REGION Network 1: จัดเก็บ
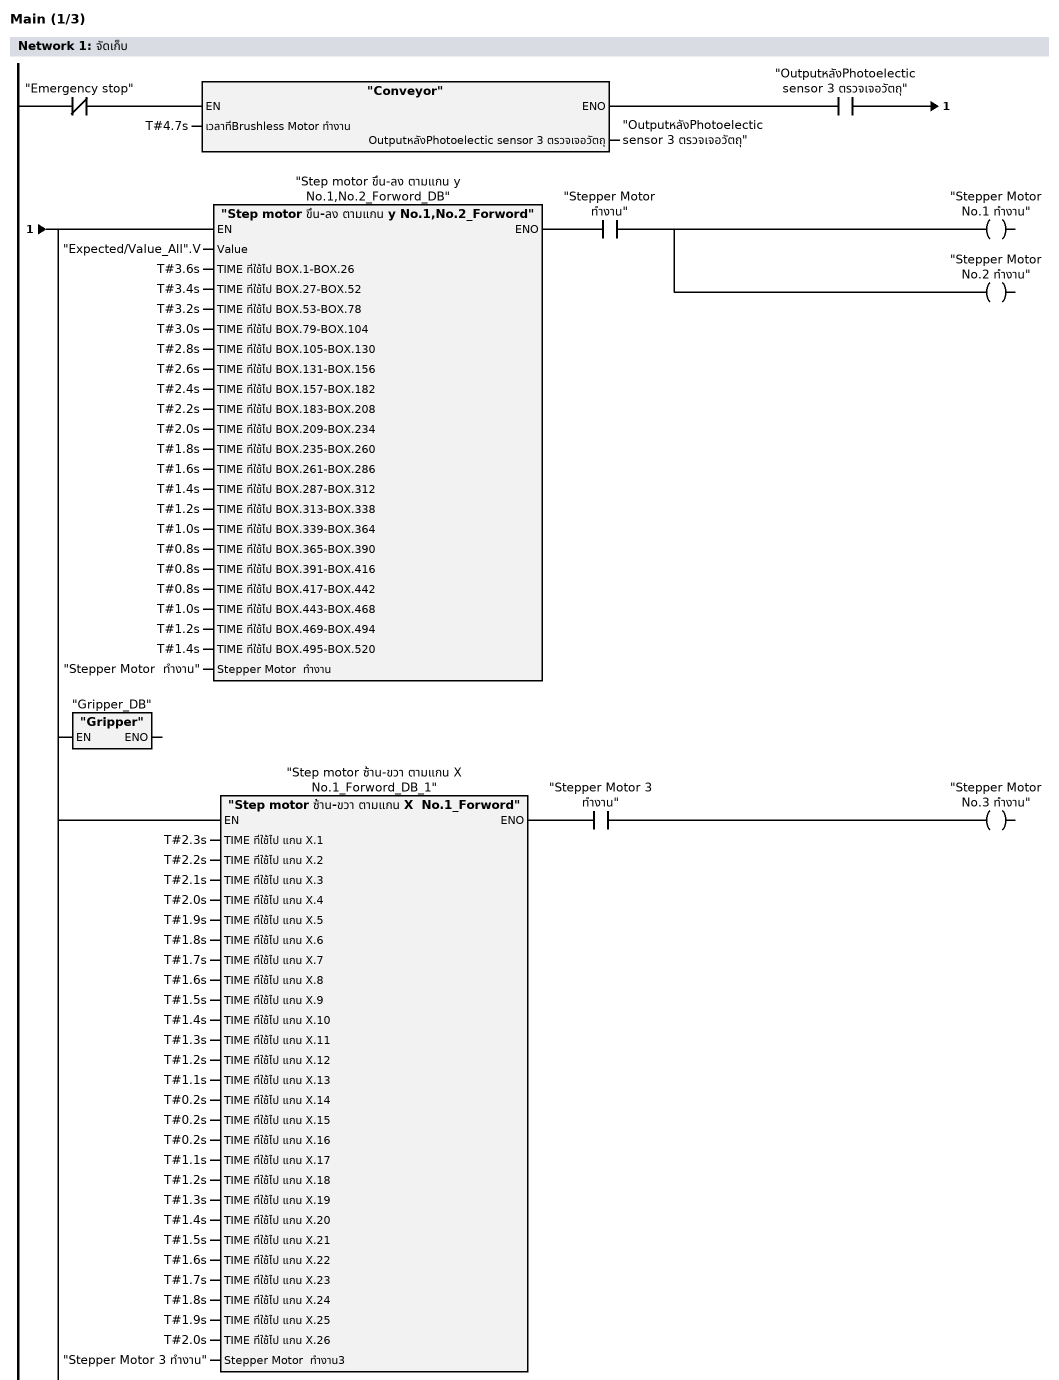
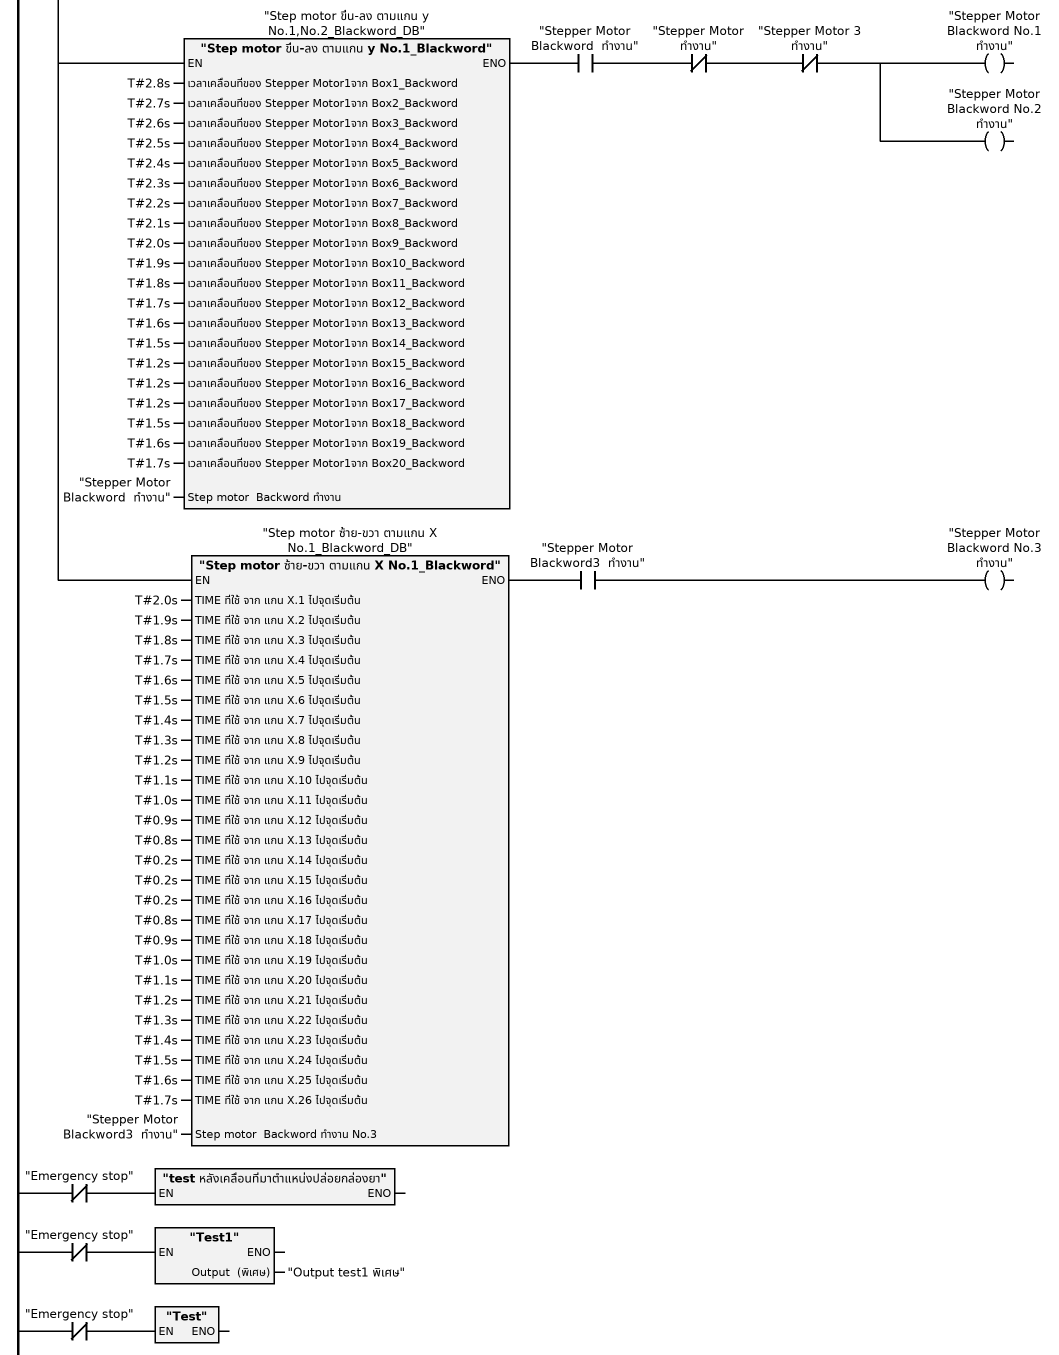
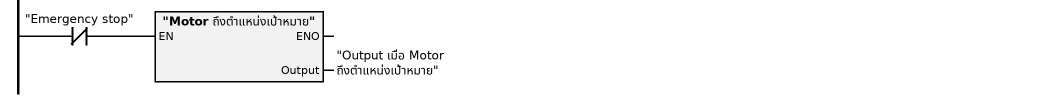
   RUNG wire#powerrail
      I_Contact( "Emergency stop" )
      "Conveyor"("เวลาที่Brushless Motor ทำงาน" := T#4.7s, "OutputหลังPhotoelectic sensor 3 ตรวจเจอวัตถุ" => "OutputหลังPhotoelectic sensor 3 ตรวจเจอวัตถุ")
      Contact( "OutputหลังPhotoelectic sensor 3 ตรวจเจอวัตถุ" )
      wire#w1
      "Step motor ขึ่น-ลง ตามแกน y No.1,No.2_Forword_DB"(Value := "Expected/Value_All".V, "TIME ที่ใช้ไป BOX.1-BOX.26" := T#3.6s, "TIME ที่ใช้ไป BOX.27-BOX.52" := T#3.4s, "TIME ที่ใช้ไป BOX.53-BOX.78" := T#3.2s, "TIME ที่ใช้ไป BOX.79-BOX.104" := T#3.0s, "TIME ที่ใช้ไป BOX.105-BOX.130" := T#2.8s, "TIME ที่ใช้ไป BOX.131-BOX.156" := T#2.6s, "TIME ที่ใช้ไป BOX.157-BOX.182" := T#2.4s, "TIME ที่ใช้ไป BOX.183-BOX.208" := T#2.2s, "TIME ที่ใช้ไป BOX.209-BOX.234" := T#2.0s, "TIME ที่ใช้ไป BOX.235-BOX.260" := T#1.8s, "TIME ที่ใช้ไป BOX.261-BOX.286" := T#1.6s, "TIME ที่ใช้ไป BOX.287-BOX.312" := T#1.4s, "TIME ที่ใช้ไป BOX.313-BOX.338" := T#1.2s, "TIME ที่ใช้ไป BOX.339-BOX.364" := T#1.0s, "TIME ที่ใช้ไป BOX.365-BOX.390" := T#0.8s, "TIME ที่ใช้ไป BOX.391-BOX.416" := T#0.8s, "TIME ที่ใช้ไป BOX.417-BOX.442" := T#0.8s, "TIME ที่ใช้ไป BOX.443-BOX.468" := T#1.0s, "TIME ที่ใช้ไป BOX.469-BOX.494" := T#1.2s, "TIME ที่ใช้ไป BOX.495-BOX.520" := T#1.4s, "Stepper Motor  ทำงาน" := "Stepper Motor  ทำงาน")
      Contact( "Stepper Motor  ทำงาน" )
      wire#w2
      Coil( "Stepper Motor No.1 ทำงาน" )
   END_RUNG
   RUNG wire#w2
      Coil( "Stepper Motor No.2 ทำงาน" )
   END_RUNG
   RUNG wire#w1
      "Gripper_DB"()
   END_RUNG
   RUNG wire#w1
      "Step motor ซ้าน-ขวา ตามแกน X  No.1_Forword_DB_1"("TIME ที่ใช้ไป แกน X.1" := T#2.3s, "TIME ที่ใช้ไป แกน X.2" := T#2.2s, "TIME ที่ใช้ไป แกน X.3" := T#2.1s, "TIME ที่ใช้ไป แกน X.4" := T#2.0s, "TIME ที่ใช้ไป แกน X.5" := T#1.9s, "TIME ที่ใช้ไป แกน X.6" := T#1.8s, "TIME ที่ใช้ไป แกน X.7" := T#1.7s, "TIME ที่ใช้ไป แกน X.8" := T#1.6s, "TIME ที่ใช้ไป แกน X.9" := T#1.5s, "TIME ที่ใช้ไป แกน X.10" := T#1.4s, "TIME ที่ใช้ไป แกน X.11" := T#1.3s, "TIME ที่ใช้ไป แกน X.12" := T#1.2s, "TIME ที่ใช้ไป แกน X.13" := T#1.1s, "TIME ที่ใช้ไป แกน X.14" := T#0.2s, "TIME ที่ใช้ไป แกน X.15" := T#0.2s, "TIME ที่ใช้ไป แกน X.16" := T#0.2s, "TIME ที่ใช้ไป แกน X.17" := T#1.1s, "TIME ที่ใช้ไป แกน X.18" := T#1.2s, "TIME ที่ใช้ไป แกน X.19" := T#1.3s, "TIME ที่ใช้ไป แกน X.20" := T#1.4s, "TIME ที่ใช้ไป แกน X.21" := T#1.5s, "TIME ที่ใช้ไป แกน X.22" := T#1.6s, "TIME ที่ใช้ไป แกน X.23" := T#1.7s, "TIME ที่ใช้ไป แกน X.24" := T#1.8s, "TIME ที่ใช้ไป แกน X.25" := T#1.9s, "TIME ที่ใช้ไป แกน X.26" := T#2.0s, "Stepper Motor  ทำงาน3" := "Stepper Motor 3 ทำงาน")
      Contact( "Stepper Motor 3 ทำงาน" )
      Coil( "Stepper Motor No.3 ทำงาน" )
   END_RUNG
   RUNG wire#w1
      "Step motor ขึ่น-ลง ตามแกน y No.1,No.2_Blackword_DB"("เวลาเคลื่อนที่ของ Stepper Motor1จาก Box1_Backword" := T#2.8s, "เวลาเคลื่อนที่ของ Stepper Motor1จาก Box2_Backword" := T#2.7s, "เวลาเคลื่อนที่ของ Stepper Motor1จาก Box3_Backword" := T#2.6s, "เวลาเคลื่อนที่ของ Stepper Motor1จาก Box4_Backword" := T#2.5s, "เวลาเคลื่อนที่ของ Stepper Motor1จาก Box5_Backword" := T#2.4s, "เวลาเคลื่อนที่ของ Stepper Motor1จาก Box6_Backword" := T#2.3s, "เวลาเคลื่อนที่ของ Stepper Motor1จาก Box7_Backword" := T#2.2s, "เวลาเคลื่อนที่ของ Stepper Motor1จาก Box8_Backword" := T#2.1s, "เวลาเคลื่อนที่ของ Stepper Motor1จาก Box9_Backword" := T#2.0s, "เวลาเคลื่อนที่ของ Stepper Motor1จาก Box10_Backword" := T#1.9s, "เวลาเคลื่อนที่ของ Stepper Motor1จาก Box11_Backword" := T#1.8s, "เวลาเคลื่อนที่ของ Stepper Motor1จาก Box12_Backword" := T#1.7s, "เวลาเคลื่อนที่ของ Stepper Motor1จาก Box13_Backword" := T#1.6s, "เวลาเคลื่อนที่ของ Stepper Motor1จาก Box14_Backword" := T#1.5s, "เวลาเคลื่อนที่ของ Stepper Motor1จาก Box15_Backword" := T#1.2s, "เวลาเคลื่อนที่ของ Stepper Motor1จาก Box16_Backword" := T#1.2s, "เวลาเคลื่อนที่ของ Stepper Motor1จาก Box17_Backword" := T#1.2s, "เวลาเคลื่อนที่ของ Stepper Motor1จาก Box18_Backword" := T#1.5s, "เวลาเคลื่อนที่ของ Stepper Motor1จาก Box19_Backword" := T#1.6s, "เวลาเคลื่อนที่ของ Stepper Motor1จาก Box20_Backword" := T#1.7s, "Step motor  Backword ทำงาน" := "Stepper Motor Blackword  ทำงาน")
      Contact( "Stepper Motor Blackword  ทำงาน" )
      I_Contact( "Stepper Motor  ทำงาน" )
      I_Contact( "Stepper Motor 3 ทำงาน" )
      wire#w3
      Coil( "Stepper Motor Blackword No.1 ทำงาน" )
   END_RUNG
   RUNG wire#w3
      Coil( "Stepper Motor Blackword No.2 ทำงาน" )
   END_RUNG
   RUNG wire#w1
      "Step motor ซ้าย-ขวา ตามแกน X No.1_Blackword_DB"("TIME ที่ใช้ จาก แกน X.1 ไปจุดเริ่มต้น" := T#2.0s, "TIME ที่ใช้ จาก แกน X.2 ไปจุดเริ่มต้น" := T#1.9s, "TIME ที่ใช้ จาก แกน X.3 ไปจุดเริ่มต้น" := T#1.8s, "TIME ที่ใช้ จาก แกน X.4 ไปจุดเริ่มต้น" := T#1.7s, "TIME ที่ใช้ จาก แกน X.5 ไปจุดเริ่มต้น" := T#1.6s, "TIME ที่ใช้ จาก แกน X.6 ไปจุดเริ่มต้น" := T#1.5s, "TIME ที่ใช้ จาก แกน X.7 ไปจุดเริ่มต้น" := T#1.4s, "TIME ที่ใช้ จาก แกน X.8 ไปจุดเริ่มต้น" := T#1.3s, "TIME ที่ใช้ จาก แกน X.9 ไปจุดเริ่มต้น" := T#1.2s, "TIME ที่ใช้ จาก แกน X.10 ไปจุดเริ่มต้น" := T#1.1s, "TIME ที่ใช้ จาก แกน X.11 ไปจุดเริ่มต้น" := T#1.0s, "TIME ที่ใช้ จาก แกน X.12 ไปจุดเริ่มต้น" := T#0.9s, "TIME ที่ใช้ จาก แกน X.13 ไปจุดเริ่มต้น" := T#0.8s, "TIME ที่ใช้ จาก แกน X.14 ไปจุดเริ่มต้น" := T#0.2s, "TIME ที่ใช้ จาก แกน X.15 ไปจุดเริ่มต้น" := T#0.2s, "TIME ที่ใช้ จาก แกน X.16 ไปจุดเริ่มต้น" := T#0.2s, "TIME ที่ใช้ จาก แกน X.17 ไปจุดเริ่มต้น" := T#0.8s, "TIME ที่ใช้ จาก แกน X.18 ไปจุดเริ่มต้น" := T#0.9s, "TIME ที่ใช้ จาก แกน X.19 ไปจุดเริ่มต้น" := T#1.0s, "TIME ที่ใช้ จาก แกน X.20 ไปจุดเริ่มต้น" := T#1.1s, "TIME ที่ใช้ จาก แกน X.21 ไปจุดเริ่มต้น" := T#1.2s, "TIME ที่ใช้ จาก แกน X.22 ไปจุดเริ่มต้น" := T#1.3s, "TIME ที่ใช้ จาก แกน X.23 ไปจุดเริ่มต้น" := T#1.4s, "TIME ที่ใช้ จาก แกน X.24 ไปจุดเริ่มต้น" := T#1.5s, "TIME ที่ใช้ จาก แกน X.25 ไปจุดเริ่มต้น" := T#1.6s, "TIME ที่ใช้ จาก แกน X.26 ไปจุดเริ่มต้น" := T#1.7s, "Step motor  Backword ทำงาน No.3" := "Stepper Motor Blackword3  ทำงาน")
      Contact( "Stepper Motor Blackword3  ทำงาน" )
      Coil( "Stepper Motor Blackword No.3 ทำงาน" )
   END_RUNG
   RUNG wire#powerrail
      I_Contact( "Emergency stop" )
      "test หลังเคลื่อนที่มาตำแหน่งปล่อยกล่องยา"()
   END_RUNG
   RUNG wire#powerrail
      I_Contact( "Emergency stop" )
      "Test1"("Output  (พิเศษ)" => "Output test1 พิเศษ")
   END_RUNG
   RUNG wire#powerrail
      I_Contact( "Emergency stop" )
      "Test"()
   END_RUNG
   RUNG wire#powerrail
      I_Contact( "Emergency stop" )
      "Motor ถึงตำแหน่งเป้าหมาย"(Output => "Output เมื่อ Motor ถึงตำแหน่งเป้าหมาย")
   END_RUNG
   // the same network as SCL:
   "Conveyor"(EN := NOT "Emergency stop",
              "เวลาที่Brushless Motor ทำงาน" := T#4.7s,
              "OutputหลังPhotoelectic sensor 3 ตรวจเจอวัตถุ" => "OutputหลังPhotoelectic sensor 3 ตรวจเจอวัตถุ",
              ENO => #_w1);
   #_w3 := #_w1 AND "OutputหลังPhotoelectic sensor 3 ตรวจเจอวัตถุ";
   "Step motor ขึ่น-ลง ตามแกน y No.1,No.2_Forword_DB"(EN := #_w1 AND "OutputหลังPhotoelectic sensor 3 ตรวจเจอวัตถุ",   // "Step motor ขึ่น-ลง ตามแกน y No.1,No.2_Forword"
                           Value := "Expected/Value_All".V,
                           "TIME ที่ใช้ไป BOX.1-BOX.26" := T#3.6s,
                           "TIME ที่ใช้ไป BOX.27-BOX.52" := T#3.4s,
                           "TIME ที่ใช้ไป BOX.53-BOX.78" := T#3.2s,
                           "TIME ที่ใช้ไป BOX.79-BOX.104" := T#3.0s,
                           "TIME ที่ใช้ไป BOX.105-BOX.130" := T#2.8s,
                           "TIME ที่ใช้ไป BOX.131-BOX.156" := T#2.6s,
                           "TIME ที่ใช้ไป BOX.157-BOX.182" := T#2.4s,
                           "TIME ที่ใช้ไป BOX.183-BOX.208" := T#2.2s,
                           "TIME ที่ใช้ไป BOX.209-BOX.234" := T#2.0s,
                           "TIME ที่ใช้ไป BOX.235-BOX.260" := T#1.8s,
                           "TIME ที่ใช้ไป BOX.261-BOX.286" := T#1.6s,
                           "TIME ที่ใช้ไป BOX.287-BOX.312" := T#1.4s,
                           "TIME ที่ใช้ไป BOX.313-BOX.338" := T#1.2s,
                           "TIME ที่ใช้ไป BOX.339-BOX.364" := T#1.0s,
                           "TIME ที่ใช้ไป BOX.365-BOX.390" := T#0.8s,
                           "TIME ที่ใช้ไป BOX.391-BOX.416" := T#0.8s,
                           "TIME ที่ใช้ไป BOX.417-BOX.442" := T#0.8s,
                           "TIME ที่ใช้ไป BOX.443-BOX.468" := T#1.0s,
                           "TIME ที่ใช้ไป BOX.469-BOX.494" := T#1.2s,
                           "TIME ที่ใช้ไป BOX.495-BOX.520" := T#1.4s,
                           "Stepper Motor  ทำงาน" := "Stepper Motor  ทำงาน",
                           ENO => #_w2);
   "Stepper Motor No.1 ทำงาน" := #_w2 AND "Stepper Motor  ทำงาน";
   "Stepper Motor No.2 ทำงาน" := "Stepper Motor No.1 ทำงาน";
   IF #_w3 THEN
       "Gripper_DB"();   // "Gripper"
   END_IF;
   "Step motor ซ้าน-ขวา ตามแกน X  No.1_Forword_DB_1"(EN := #_w3,   // "Step motor ซ้าน-ขวา ตามแกน X  No.1_Forword"
                           "TIME ที่ใช้ไป แกน X.1" := T#2.3s,
                           "TIME ที่ใช้ไป แกน X.2" := T#2.2s,
                           "TIME ที่ใช้ไป แกน X.3" := T#2.1s,
                           "TIME ที่ใช้ไป แกน X.4" := T#2.0s,
                           "TIME ที่ใช้ไป แกน X.5" := T#1.9s,
                           "TIME ที่ใช้ไป แกน X.6" := T#1.8s,
                           "TIME ที่ใช้ไป แกน X.7" := T#1.7s,
                           "TIME ที่ใช้ไป แกน X.8" := T#1.6s,
                           "TIME ที่ใช้ไป แกน X.9" := T#1.5s,
                           "TIME ที่ใช้ไป แกน X.10" := T#1.4s,
                           "TIME ที่ใช้ไป แกน X.11" := T#1.3s,
                           "TIME ที่ใช้ไป แกน X.12" := T#1.2s,
                           "TIME ที่ใช้ไป แกน X.13" := T#1.1s,
                           "TIME ที่ใช้ไป แกน X.14" := T#0.2s,
                           "TIME ที่ใช้ไป แกน X.15" := T#0.2s,
                           "TIME ที่ใช้ไป แกน X.16" := T#0.2s,
                           "TIME ที่ใช้ไป แกน X.17" := T#1.1s,
                           "TIME ที่ใช้ไป แกน X.18" := T#1.2s,
                           "TIME ที่ใช้ไป แกน X.19" := T#1.3s,
                           "TIME ที่ใช้ไป แกน X.20" := T#1.4s,
                           "TIME ที่ใช้ไป แกน X.21" := T#1.5s,
                           "TIME ที่ใช้ไป แกน X.22" := T#1.6s,
                           "TIME ที่ใช้ไป แกน X.23" := T#1.7s,
                           "TIME ที่ใช้ไป แกน X.24" := T#1.8s,
                           "TIME ที่ใช้ไป แกน X.25" := T#1.9s,
                           "TIME ที่ใช้ไป แกน X.26" := T#2.0s,
                           "Stepper Motor  ทำงาน3" := "Stepper Motor 3 ทำงาน",
                           ENO => #_w4);
   "Stepper Motor No.3 ทำงาน" := #_w4 AND "Stepper Motor 3 ทำงาน";
   "Step motor ขึ่น-ลง ตามแกน y No.1,No.2_Blackword_DB"(EN := #_w3,   // "Step motor ขึ่น-ลง ตามแกน y No.1_Blackword"
                           "เวลาเคลื่อนที่ของ Stepper Motor1จาก Box1_Backword" := T#2.8s,
                           "เวลาเคลื่อนที่ของ Stepper Motor1จาก Box2_Backword" := T#2.7s,
                           "เวลาเคลื่อนที่ของ Stepper Motor1จาก Box3_Backword" := T#2.6s,
                           "เวลาเคลื่อนที่ของ Stepper Motor1จาก Box4_Backword" := T#2.5s,
                           "เวลาเคลื่อนที่ของ Stepper Motor1จาก Box5_Backword" := T#2.4s,
                           "เวลาเคลื่อนที่ของ Stepper Motor1จาก Box6_Backword" := T#2.3s,
                           "เวลาเคลื่อนที่ของ Stepper Motor1จาก Box7_Backword" := T#2.2s,
                           "เวลาเคลื่อนที่ของ Stepper Motor1จาก Box8_Backword" := T#2.1s,
                           "เวลาเคลื่อนที่ของ Stepper Motor1จาก Box9_Backword" := T#2.0s,
                           "เวลาเคลื่อนที่ของ Stepper Motor1จาก Box10_Backword" := T#1.9s,
                           "เวลาเคลื่อนที่ของ Stepper Motor1จาก Box11_Backword" := T#1.8s,
                           "เวลาเคลื่อนที่ของ Stepper Motor1จาก Box12_Backword" := T#1.7s,
                           "เวลาเคลื่อนที่ของ Stepper Motor1จาก Box13_Backword" := T#1.6s,
                           "เวลาเคลื่อนที่ของ Stepper Motor1จาก Box14_Backword" := T#1.5s,
                           "เวลาเคลื่อนที่ของ Stepper Motor1จาก Box15_Backword" := T#1.2s,
                           "เวลาเคลื่อนที่ของ Stepper Motor1จาก Box16_Backword" := T#1.2s,
                           "เวลาเคลื่อนที่ของ Stepper Motor1จาก Box17_Backword" := T#1.2s,
                           "เวลาเคลื่อนที่ของ Stepper Motor1จาก Box18_Backword" := T#1.5s,
                           "เวลาเคลื่อนที่ของ Stepper Motor1จาก Box19_Backword" := T#1.6s,
                           "เวลาเคลื่อนที่ของ Stepper Motor1จาก Box20_Backword" := T#1.7s,
                           "Step motor  Backword ทำงาน" := "Stepper Motor Blackword  ทำงาน",
                           ENO => #_w5);
   "Stepper Motor Blackword No.1 ทำงาน" := #_w5 AND "Stepper Motor Blackword  ทำงาน" AND NOT "Stepper Motor  ทำงาน" AND NOT "Stepper Motor 3 ทำงาน";
   "Stepper Motor Blackword No.2 ทำงาน" := "Stepper Motor Blackword No.1 ทำงาน";
   "Step motor ซ้าย-ขวา ตามแกน X No.1_Blackword_DB"(EN := #_w3,   // "Step motor ซ้าย-ขวา ตามแกน X No.1_Blackword"
                           "TIME ที่ใช้ จาก แกน X.1 ไปจุดเริ่มต้น" := T#2.0s,
                           "TIME ที่ใช้ จาก แกน X.2 ไปจุดเริ่มต้น" := T#1.9s,
                           "TIME ที่ใช้ จาก แกน X.3 ไปจุดเริ่มต้น" := T#1.8s,
                           "TIME ที่ใช้ จาก แกน X.4 ไปจุดเริ่มต้น" := T#1.7s,
                           "TIME ที่ใช้ จาก แกน X.5 ไปจุดเริ่มต้น" := T#1.6s,
                           "TIME ที่ใช้ จาก แกน X.6 ไปจุดเริ่มต้น" := T#1.5s,
                           "TIME ที่ใช้ จาก แกน X.7 ไปจุดเริ่มต้น" := T#1.4s,
                           "TIME ที่ใช้ จาก แกน X.8 ไปจุดเริ่มต้น" := T#1.3s,
                           "TIME ที่ใช้ จาก แกน X.9 ไปจุดเริ่มต้น" := T#1.2s,
                           "TIME ที่ใช้ จาก แกน X.10 ไปจุดเริ่มต้น" := T#1.1s,
                           "TIME ที่ใช้ จาก แกน X.11 ไปจุดเริ่มต้น" := T#1.0s,
                           "TIME ที่ใช้ จาก แกน X.12 ไปจุดเริ่มต้น" := T#0.9s,
                           "TIME ที่ใช้ จาก แกน X.13 ไปจุดเริ่มต้น" := T#0.8s,
                           "TIME ที่ใช้ จาก แกน X.14 ไปจุดเริ่มต้น" := T#0.2s,
                           "TIME ที่ใช้ จาก แกน X.15 ไปจุดเริ่มต้น" := T#0.2s,
                           "TIME ที่ใช้ จาก แกน X.16 ไปจุดเริ่มต้น" := T#0.2s,
                           "TIME ที่ใช้ จาก แกน X.17 ไปจุดเริ่มต้น" := T#0.8s,
                           "TIME ที่ใช้ จาก แกน X.18 ไปจุดเริ่มต้น" := T#0.9s,
                           "TIME ที่ใช้ จาก แกน X.19 ไปจุดเริ่มต้น" := T#1.0s,
                           "TIME ที่ใช้ จาก แกน X.20 ไปจุดเริ่มต้น" := T#1.1s,
                           "TIME ที่ใช้ จาก แกน X.21 ไปจุดเริ่มต้น" := T#1.2s,
                           "TIME ที่ใช้ จาก แกน X.22 ไปจุดเริ่มต้น" := T#1.3s,
                           "TIME ที่ใช้ จาก แกน X.23 ไปจุดเริ่มต้น" := T#1.4s,
                           "TIME ที่ใช้ จาก แกน X.24 ไปจุดเริ่มต้น" := T#1.5s,
                           "TIME ที่ใช้ จาก แกน X.25 ไปจุดเริ่มต้น" := T#1.6s,
                           "TIME ที่ใช้ จาก แกน X.26 ไปจุดเริ่มต้น" := T#1.7s,
                           "Step motor  Backword ทำงาน No.3" := "Stepper Motor Blackword3  ทำงาน",
                           ENO => #_w6);
   "Stepper Motor Blackword No.3 ทำงาน" := #_w6 AND "Stepper Motor Blackword3  ทำงาน";
   IF NOT "Emergency stop" THEN "test หลังเคลื่อนที่มาตำแหน่งปล่อยกล่องยา"(); END_IF;
   IF NOT "Emergency stop" THEN "Test1"("Output  (พิเศษ)" => "Output test1 พิเศษ"); END_IF;
   IF NOT "Emergency stop" THEN "Test"(); END_IF;
   IF NOT "Emergency stop" THEN
       "Motor ถึงตำแหน่งเป้าหมาย"(Output => "Output เมื่อ Motor ถึงตำแหน่งเป้าหมาย");
   END_IF;
END_REGION

REGION Network 2: เบิกจ่าย
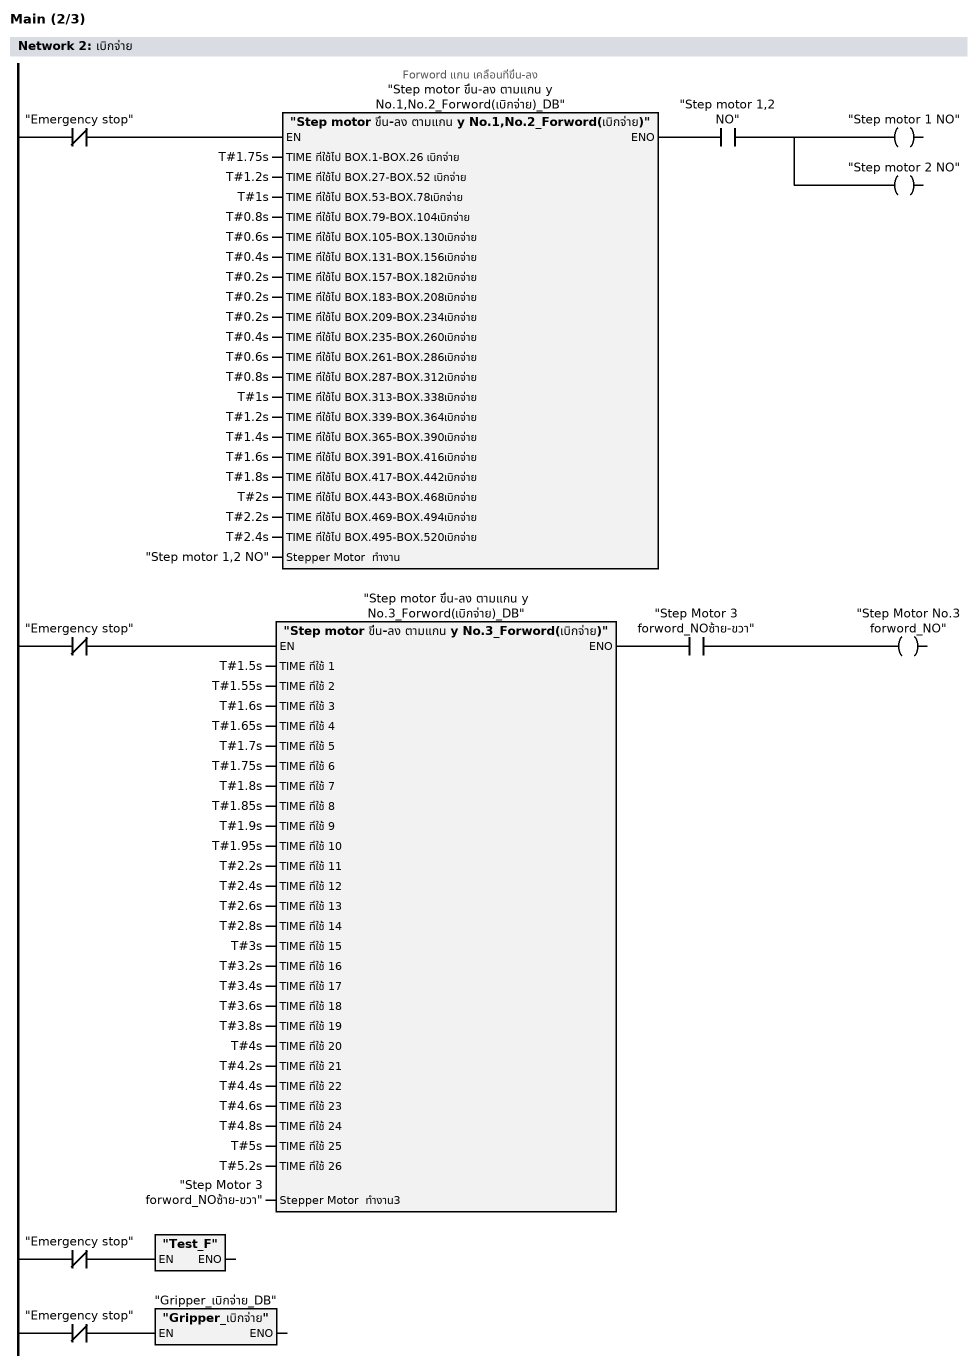
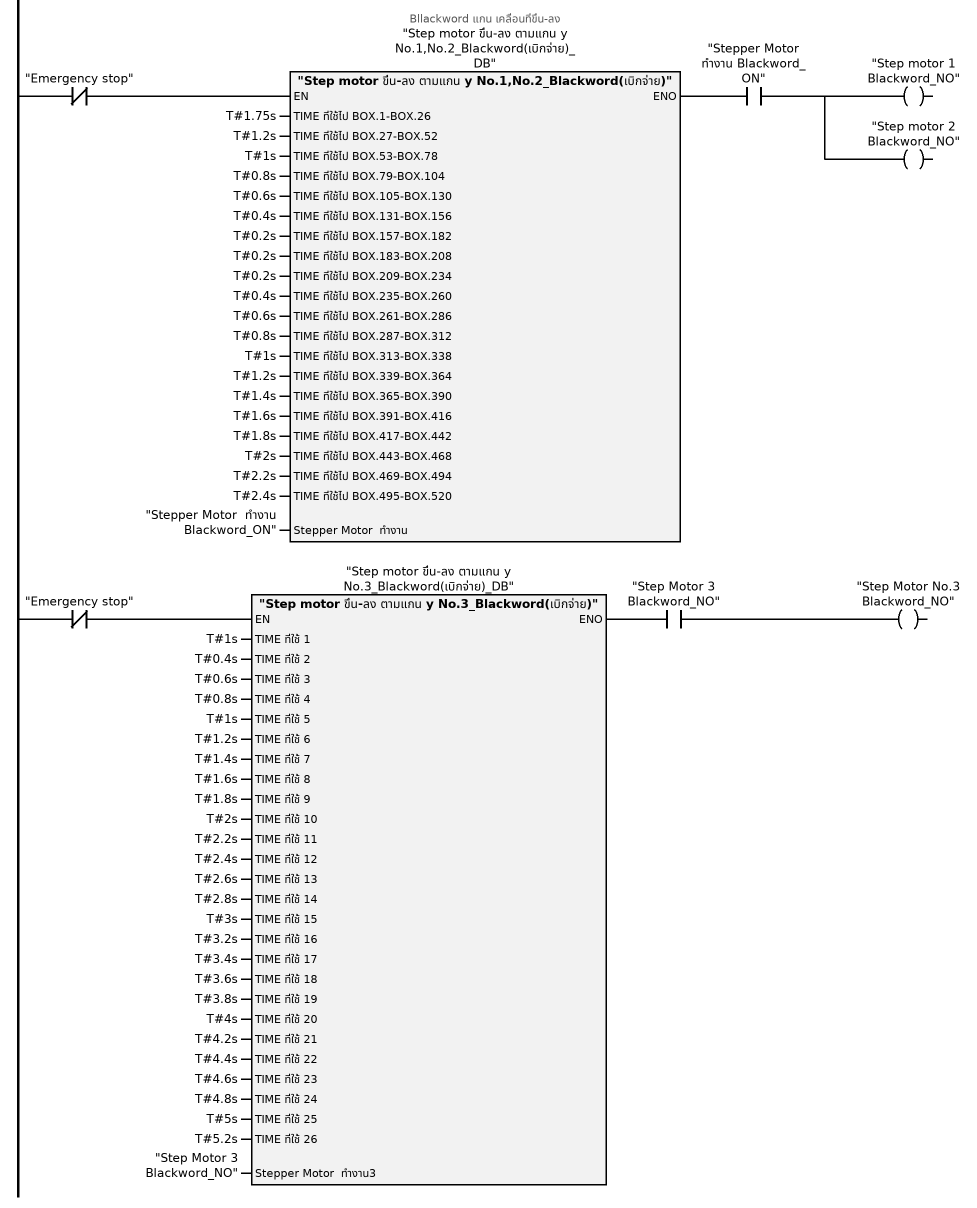
   RUNG wire#powerrail
      I_Contact( "Emergency stop" )
      "Step motor ขึ่น-ลง ตามแกน y No.1,No.2_Forword(เบิกจ่าย)_DB"("TIME ที่ใช้ไป BOX.1-BOX.26 เบิกจ่าย" := T#1.75s, "TIME ที่ใช้ไป BOX.27-BOX.52 เบิกจ่าย" := T#1.2s, "TIME ที่ใช้ไป BOX.53-BOX.78เบิกจ่าย" := T#1s, "TIME ที่ใช้ไป BOX.79-BOX.104เบิกจ่าย" := T#0.8s, "TIME ที่ใช้ไป BOX.105-BOX.130เบิกจ่าย" := T#0.6s, "TIME ที่ใช้ไป BOX.131-BOX.156เบิกจ่าย" := T#0.4s, "TIME ที่ใช้ไป BOX.157-BOX.182เบิกจ่าย" := T#0.2s, "TIME ที่ใช้ไป BOX.183-BOX.208เบิกจ่าย" := T#0.2s, "TIME ที่ใช้ไป BOX.209-BOX.234เบิกจ่าย" := T#0.2s, "TIME ที่ใช้ไป BOX.235-BOX.260เบิกจ่าย" := T#0.4s, "TIME ที่ใช้ไป BOX.261-BOX.286เบิกจ่าย" := T#0.6s, "TIME ที่ใช้ไป BOX.287-BOX.312เบิกจ่าย" := T#0.8s, "TIME ที่ใช้ไป BOX.313-BOX.338เบิกจ่าย" := T#1s, "TIME ที่ใช้ไป BOX.339-BOX.364เบิกจ่าย" := T#1.2s, "TIME ที่ใช้ไป BOX.365-BOX.390เบิกจ่าย" := T#1.4s, "TIME ที่ใช้ไป BOX.391-BOX.416เบิกจ่าย" := T#1.6s, "TIME ที่ใช้ไป BOX.417-BOX.442เบิกจ่าย" := T#1.8s, "TIME ที่ใช้ไป BOX.443-BOX.468เบิกจ่าย" := T#2s, "TIME ที่ใช้ไป BOX.469-BOX.494เบิกจ่าย" := T#2.2s, "TIME ที่ใช้ไป BOX.495-BOX.520เบิกจ่าย" := T#2.4s, "Stepper Motor  ทำงาน" := "Step motor 1,2 NO")   // Forword แกน เคลื่อนที่ขึ่น-ลง
      Contact( "Step motor 1,2 NO" )
      wire#w1
      Coil( "Step motor 1 NO" )
   END_RUNG
   RUNG wire#w1
      Coil( "Step motor 2 NO" )
   END_RUNG
   RUNG wire#powerrail
      I_Contact( "Emergency stop" )
      "Step motor ขึ่น-ลง ตามแกน y No.3_Forword(เบิกจ่าย)_DB"("TIME ที่ใช้ 1" := T#1.5s, "TIME ที่ใช้ 2" := T#1.55s, "TIME ที่ใช้ 3" := T#1.6s, "TIME ที่ใช้ 4" := T#1.65s, "TIME ที่ใช้ 5" := T#1.7s, "TIME ที่ใช้ 6" := T#1.75s, "TIME ที่ใช้ 7" := T#1.8s, "TIME ที่ใช้ 8" := T#1.85s, "TIME ที่ใช้ 9" := T#1.9s, "TIME ที่ใช้ 10" := T#1.95s, "TIME ที่ใช้ 11" := T#2.2s, "TIME ที่ใช้ 12" := T#2.4s, "TIME ที่ใช้ 13" := T#2.6s, "TIME ที่ใช้ 14" := T#2.8s, "TIME ที่ใช้ 15" := T#3s, "TIME ที่ใช้ 16" := T#3.2s, "TIME ที่ใช้ 17" := T#3.4s, "TIME ที่ใช้ 18" := T#3.6s, "TIME ที่ใช้ 19" := T#3.8s, "TIME ที่ใช้ 20" := T#4s, "TIME ที่ใช้ 21" := T#4.2s, "TIME ที่ใช้ 22" := T#4.4s, "TIME ที่ใช้ 23" := T#4.6s, "TIME ที่ใช้ 24" := T#4.8s, "TIME ที่ใช้ 25" := T#5s, "TIME ที่ใช้ 26" := T#5.2s, "Stepper Motor  ทำงาน3" := "Step Motor 3 forword_NOซ้าย-ขวา")
      Contact( "Step Motor 3 forword_NOซ้าย-ขวา" )
      Coil( "Step Motor No.3 forword_NO" )
   END_RUNG
   RUNG wire#powerrail
      I_Contact( "Emergency stop" )
      "Test_F"()
   END_RUNG
   RUNG wire#powerrail
      I_Contact( "Emergency stop" )
      "Gripper_เบิกจ่าย_DB"()
   END_RUNG
   RUNG wire#powerrail
      I_Contact( "Emergency stop" )
      "Step motor ขึ่น-ลง ตามแกน y No.1,No.2_Blackword(เบิกจ่าย)_DB"("TIME ที่ใช้ไป BOX.1-BOX.26" := T#1.75s, "TIME ที่ใช้ไป BOX.27-BOX.52" := T#1.2s, "TIME ที่ใช้ไป BOX.53-BOX.78" := T#1s, "TIME ที่ใช้ไป BOX.79-BOX.104" := T#0.8s, "TIME ที่ใช้ไป BOX.105-BOX.130" := T#0.6s, "TIME ที่ใช้ไป BOX.131-BOX.156" := T#0.4s, "TIME ที่ใช้ไป BOX.157-BOX.182" := T#0.2s, "TIME ที่ใช้ไป BOX.183-BOX.208" := T#0.2s, "TIME ที่ใช้ไป BOX.209-BOX.234" := T#0.2s, "TIME ที่ใช้ไป BOX.235-BOX.260" := T#0.4s, "TIME ที่ใช้ไป BOX.261-BOX.286" := T#0.6s, "TIME ที่ใช้ไป BOX.287-BOX.312" := T#0.8s, "TIME ที่ใช้ไป BOX.313-BOX.338" := T#1s, "TIME ที่ใช้ไป BOX.339-BOX.364" := T#1.2s, "TIME ที่ใช้ไป BOX.365-BOX.390" := T#1.4s, "TIME ที่ใช้ไป BOX.391-BOX.416" := T#1.6s, "TIME ที่ใช้ไป BOX.417-BOX.442" := T#1.8s, "TIME ที่ใช้ไป BOX.443-BOX.468" := T#2s, "TIME ที่ใช้ไป BOX.469-BOX.494" := T#2.2s, "TIME ที่ใช้ไป BOX.495-BOX.520" := T#2.4s, "Stepper Motor  ทำงาน" := "Stepper Motor  ทำงาน Blackword_ON")   // Bllackword แกน เคลื่อนที่ขึ่น-ลง
      Contact( "Stepper Motor  ทำงาน Blackword_ON" )
      wire#w2
      Coil( "Step motor 1 Blackword_NO" )
   END_RUNG
   RUNG wire#w2
      Coil( "Step motor 2 Blackword_NO" )
   END_RUNG
   RUNG wire#powerrail
      I_Contact( "Emergency stop" )
      "Step motor ขึ่น-ลง ตามแกน y No.3_Blackword(เบิกจ่าย)_DB"("TIME ที่ใช้ 1" := T#1s, "TIME ที่ใช้ 2" := T#0.4s, "TIME ที่ใช้ 3" := T#0.6s, "TIME ที่ใช้ 4" := T#0.8s, "TIME ที่ใช้ 5" := T#1s, "TIME ที่ใช้ 6" := T#1.2s, "TIME ที่ใช้ 7" := T#1.4s, "TIME ที่ใช้ 8" := T#1.6s, "TIME ที่ใช้ 9" := T#1.8s, "TIME ที่ใช้ 10" := T#2s, "TIME ที่ใช้ 11" := T#2.2s, "TIME ที่ใช้ 12" := T#2.4s, "TIME ที่ใช้ 13" := T#2.6s, "TIME ที่ใช้ 14" := T#2.8s, "TIME ที่ใช้ 15" := T#3s, "TIME ที่ใช้ 16" := T#3.2s, "TIME ที่ใช้ 17" := T#3.4s, "TIME ที่ใช้ 18" := T#3.6s, "TIME ที่ใช้ 19" := T#3.8s, "TIME ที่ใช้ 20" := T#4s, "TIME ที่ใช้ 21" := T#4.2s, "TIME ที่ใช้ 22" := T#4.4s, "TIME ที่ใช้ 23" := T#4.6s, "TIME ที่ใช้ 24" := T#4.8s, "TIME ที่ใช้ 25" := T#5s, "TIME ที่ใช้ 26" := T#5.2s, "Stepper Motor  ทำงาน3" := "Step Motor 3 Blackword_NO")
      Contact( "Step Motor 3 Blackword_NO" )
      Coil( "Step Motor No.3 Blackword_NO" )
   END_RUNG
   // the same network as SCL:
   "Step motor ขึ่น-ลง ตามแกน y No.1,No.2_Forword(เบิกจ่าย)_DB"(EN := NOT "Emergency stop",   // "Step motor ขึ่น-ลง ตามแกน y No.1,No.2_Forword(เบิกจ่าย)": Forword แกน เคลื่อนที่ขึ่น-ลง
                           "TIME ที่ใช้ไป BOX.1-BOX.26 เบิกจ่าย" := T#1.75s,
                           "TIME ที่ใช้ไป BOX.27-BOX.52 เบิกจ่าย" := T#1.2s,
                           "TIME ที่ใช้ไป BOX.53-BOX.78เบิกจ่าย" := T#1s,
                           "TIME ที่ใช้ไป BOX.79-BOX.104เบิกจ่าย" := T#0.8s,
                           "TIME ที่ใช้ไป BOX.105-BOX.130เบิกจ่าย" := T#0.6s,
                           "TIME ที่ใช้ไป BOX.131-BOX.156เบิกจ่าย" := T#0.4s,
                           "TIME ที่ใช้ไป BOX.157-BOX.182เบิกจ่าย" := T#0.2s,
                           "TIME ที่ใช้ไป BOX.183-BOX.208เบิกจ่าย" := T#0.2s,
                           "TIME ที่ใช้ไป BOX.209-BOX.234เบิกจ่าย" := T#0.2s,
                           "TIME ที่ใช้ไป BOX.235-BOX.260เบิกจ่าย" := T#0.4s,
                           "TIME ที่ใช้ไป BOX.261-BOX.286เบิกจ่าย" := T#0.6s,
                           "TIME ที่ใช้ไป BOX.287-BOX.312เบิกจ่าย" := T#0.8s,
                           "TIME ที่ใช้ไป BOX.313-BOX.338เบิกจ่าย" := T#1s,
                           "TIME ที่ใช้ไป BOX.339-BOX.364เบิกจ่าย" := T#1.2s,
                           "TIME ที่ใช้ไป BOX.365-BOX.390เบิกจ่าย" := T#1.4s,
                           "TIME ที่ใช้ไป BOX.391-BOX.416เบิกจ่าย" := T#1.6s,
                           "TIME ที่ใช้ไป BOX.417-BOX.442เบิกจ่าย" := T#1.8s,
                           "TIME ที่ใช้ไป BOX.443-BOX.468เบิกจ่าย" := T#2s,
                           "TIME ที่ใช้ไป BOX.469-BOX.494เบิกจ่าย" := T#2.2s,
                           "TIME ที่ใช้ไป BOX.495-BOX.520เบิกจ่าย" := T#2.4s,
                           "Stepper Motor  ทำงาน" := "Step motor 1,2 NO",
                           ENO => #_w1);
   "Step motor 1 NO" := #_w1 AND "Step motor 1,2 NO";
   "Step motor 2 NO" := "Step motor 1 NO";
   "Step motor ขึ่น-ลง ตามแกน y No.3_Forword(เบิกจ่าย)_DB"(EN := NOT "Emergency stop",   // "Step motor ขึ่น-ลง ตามแกน y No.3_Forword(เบิกจ่าย)"
                           "TIME ที่ใช้ 1" := T#1.5s,
                           "TIME ที่ใช้ 2" := T#1.55s,
                           "TIME ที่ใช้ 3" := T#1.6s,
                           "TIME ที่ใช้ 4" := T#1.65s,
                           "TIME ที่ใช้ 5" := T#1.7s,
                           "TIME ที่ใช้ 6" := T#1.75s,
                           "TIME ที่ใช้ 7" := T#1.8s,
                           "TIME ที่ใช้ 8" := T#1.85s,
                           "TIME ที่ใช้ 9" := T#1.9s,
                           "TIME ที่ใช้ 10" := T#1.95s,
                           "TIME ที่ใช้ 11" := T#2.2s,
                           "TIME ที่ใช้ 12" := T#2.4s,
                           "TIME ที่ใช้ 13" := T#2.6s,
                           "TIME ที่ใช้ 14" := T#2.8s,
                           "TIME ที่ใช้ 15" := T#3s,
                           "TIME ที่ใช้ 16" := T#3.2s,
                           "TIME ที่ใช้ 17" := T#3.4s,
                           "TIME ที่ใช้ 18" := T#3.6s,
                           "TIME ที่ใช้ 19" := T#3.8s,
                           "TIME ที่ใช้ 20" := T#4s,
                           "TIME ที่ใช้ 21" := T#4.2s,
                           "TIME ที่ใช้ 22" := T#4.4s,
                           "TIME ที่ใช้ 23" := T#4.6s,
                           "TIME ที่ใช้ 24" := T#4.8s,
                           "TIME ที่ใช้ 25" := T#5s,
                           "TIME ที่ใช้ 26" := T#5.2s,
                           "Stepper Motor  ทำงาน3" := "Step Motor 3 forword_NOซ้าย-ขวา",
                           ENO => #_w2);
   "Step Motor No.3 forword_NO" := #_w2 AND "Step Motor 3 forword_NOซ้าย-ขวา";
   IF NOT "Emergency stop" THEN "Test_F"(); END_IF;
   IF NOT "Emergency stop" THEN
       "Gripper_เบิกจ่าย_DB"();   // "Gripper_เบิกจ่าย"
   END_IF;
   "Step motor ขึ่น-ลง ตามแกน y No.1,No.2_Blackword(เบิกจ่าย)_DB"(EN := NOT "Emergency stop",   // "Step motor ขึ่น-ลง ตามแกน y No.1,No.2_Blackword(เบิกจ่าย)": Bllackword แกน เคลื่อนที่ขึ่น-ลง
                           "TIME ที่ใช้ไป BOX.1-BOX.26" := T#1.75s,
                           "TIME ที่ใช้ไป BOX.27-BOX.52" := T#1.2s,
                           "TIME ที่ใช้ไป BOX.53-BOX.78" := T#1s,
                           "TIME ที่ใช้ไป BOX.79-BOX.104" := T#0.8s,
                           "TIME ที่ใช้ไป BOX.105-BOX.130" := T#0.6s,
                           "TIME ที่ใช้ไป BOX.131-BOX.156" := T#0.4s,
                           "TIME ที่ใช้ไป BOX.157-BOX.182" := T#0.2s,
                           "TIME ที่ใช้ไป BOX.183-BOX.208" := T#0.2s,
                           "TIME ที่ใช้ไป BOX.209-BOX.234" := T#0.2s,
                           "TIME ที่ใช้ไป BOX.235-BOX.260" := T#0.4s,
                           "TIME ที่ใช้ไป BOX.261-BOX.286" := T#0.6s,
                           "TIME ที่ใช้ไป BOX.287-BOX.312" := T#0.8s,
                           "TIME ที่ใช้ไป BOX.313-BOX.338" := T#1s,
                           "TIME ที่ใช้ไป BOX.339-BOX.364" := T#1.2s,
                           "TIME ที่ใช้ไป BOX.365-BOX.390" := T#1.4s,
                           "TIME ที่ใช้ไป BOX.391-BOX.416" := T#1.6s,
                           "TIME ที่ใช้ไป BOX.417-BOX.442" := T#1.8s,
                           "TIME ที่ใช้ไป BOX.443-BOX.468" := T#2s,
                           "TIME ที่ใช้ไป BOX.469-BOX.494" := T#2.2s,
                           "TIME ที่ใช้ไป BOX.495-BOX.520" := T#2.4s,
                           "Stepper Motor  ทำงาน" := "Stepper Motor  ทำงาน Blackword_ON",
                           ENO => #_w3);
   "Step motor 1 Blackword_NO" := #_w3 AND "Stepper Motor  ทำงาน Blackword_ON";
   "Step motor 2 Blackword_NO" := "Step motor 1 Blackword_NO";
   "Step motor ขึ่น-ลง ตามแกน y No.3_Blackword(เบิกจ่าย)_DB"(EN := NOT "Emergency stop",   // "Step motor ขึ่น-ลง ตามแกน y No.3_Blackword(เบิกจ่าย)"
                           "TIME ที่ใช้ 1" := T#1s,
                           "TIME ที่ใช้ 2" := T#0.4s,
                           "TIME ที่ใช้ 3" := T#0.6s,
                           "TIME ที่ใช้ 4" := T#0.8s,
                           "TIME ที่ใช้ 5" := T#1s,
                           "TIME ที่ใช้ 6" := T#1.2s,
                           "TIME ที่ใช้ 7" := T#1.4s,
                           "TIME ที่ใช้ 8" := T#1.6s,
                           "TIME ที่ใช้ 9" := T#1.8s,
                           "TIME ที่ใช้ 10" := T#2s,
                           "TIME ที่ใช้ 11" := T#2.2s,
                           "TIME ที่ใช้ 12" := T#2.4s,
                           "TIME ที่ใช้ 13" := T#2.6s,
                           "TIME ที่ใช้ 14" := T#2.8s,
                           "TIME ที่ใช้ 15" := T#3s,
                           "TIME ที่ใช้ 16" := T#3.2s,
                           "TIME ที่ใช้ 17" := T#3.4s,
                           "TIME ที่ใช้ 18" := T#3.6s,
                           "TIME ที่ใช้ 19" := T#3.8s,
                           "TIME ที่ใช้ 20" := T#4s,
                           "TIME ที่ใช้ 21" := T#4.2s,
                           "TIME ที่ใช้ 22" := T#4.4s,
                           "TIME ที่ใช้ 23" := T#4.6s,
                           "TIME ที่ใช้ 24" := T#4.8s,
                           "TIME ที่ใช้ 25" := T#5s,
                           "TIME ที่ใช้ 26" := T#5.2s,
                           "Stepper Motor  ทำงาน3" := "Step Motor 3 Blackword_NO",
                           ENO => #_w4);
   "Step Motor No.3 Blackword_NO" := #_w4 AND "Step Motor 3 Blackword_NO";
END_REGION

REGION Network 3: Screen
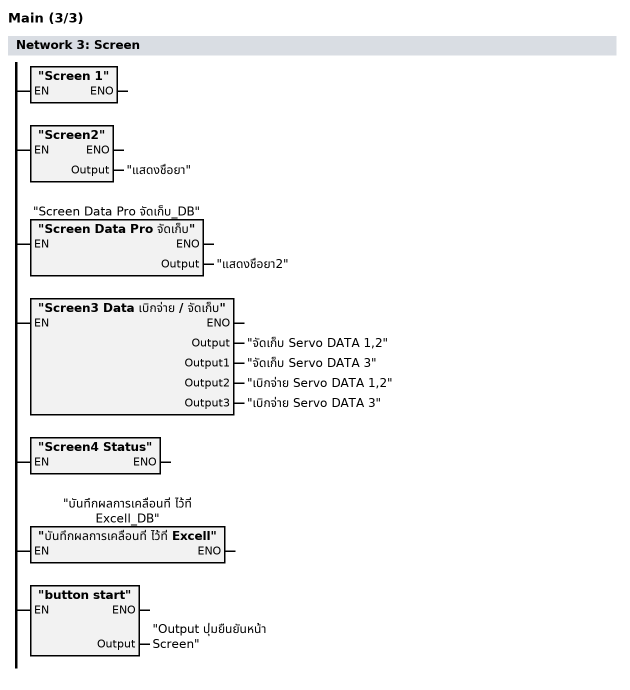
   RUNG wire#powerrail
      "Screen 1"()
   END_RUNG
   RUNG wire#powerrail
      "Screen2"(Output => "แสดงชื่อยา")
   END_RUNG
   RUNG wire#powerrail
      "Screen Data Pro จัดเก็บ_DB"(Output => "แสดงชื่อยา2")
   END_RUNG
   RUNG wire#powerrail
      "Screen3 Data เบิกจ่าย / จัดเก็บ"(Output => "จัดเก็บ Servo DATA 1,2", Output1 => "จัดเก็บ Servo DATA 3", Output2 => "เบิกจ่าย Servo DATA 1,2", Output3 => "เบิกจ่าย Servo DATA 3")
   END_RUNG
   RUNG wire#powerrail
      "Screen4 Status"()
   END_RUNG
   RUNG wire#powerrail
      "บันทึกผลการเคลื่อนที่ ไว้ที่ Excell_DB"()
   END_RUNG
   RUNG wire#powerrail
      "button start"(Output => "Output ปุ่มยืนยันหน้า Screen")
   END_RUNG
   // the same network as SCL:
   "Screen 1"();
   "Screen2"(Output => "แสดงชื่อยา");
   "Screen Data Pro จัดเก็บ_DB"(Output => "แสดงชื่อยา2");   // "Screen Data Pro จัดเก็บ"
   "Screen3 Data เบิกจ่าย / จัดเก็บ"(Output => "จัดเก็บ Servo DATA 1,2",
                           Output1 => "จัดเก็บ Servo DATA 3",
                           Output2 => "เบิกจ่าย Servo DATA 1,2",
                           Output3 => "เบิกจ่าย Servo DATA 3");
   "Screen4 Status"();
   "บันทึกผลการเคลื่อนที่ ไว้ที่ Excell_DB"();   // "บันทึกผลการเคลื่อนที่ ไว้ที่ Excell"
   "button start"(Output => "Output ปุ่มยืนยันหน้า Screen");
END_REGION
END_ORGANIZATION_BLOCK

// folder: GRAPH

FUNCTION_BLOCK "GRAPH_จัดเก็บ"   // FB17, GRAPH_PLUS
{ S7_Optimized_Access := 'TRUE' }
VERSION : 0.1
   VAR_INPUT
      OFF_SQ : Bool := false;   // Turn sequence off
      INIT_SQ : Bool := false;   // Set sequence to initial state
      ACK_EF : Bool := false;   // Acknowledge all errors and faults
      S_PREV : Bool := false;   // Output previous step in parameter S_NO
      S_NEXT : Bool := false;   // Indicate next step in parameter S_NO
      SW_AUTO : Bool := false;   // Automatic mode
      SW_TAP : Bool := false;   // Semiautomatic/switch with transition
      SW_TOP : Bool := false;   // Semiautomatic/ignore transition
      SW_MAN : Bool := false;   // Manual mode
      S_SEL : Int := 0;   // Select step to be output to S_NO
      S_ON : Bool := false;   // Activate step indicated in S_NO
      S_OFF : Bool := false;   // Deactivate step indicated S_NO
      T_PUSH : Bool := false;   // Enable transition to switch in semi automatic mode
   END_VAR
   VAR_OUTPUT
      S_NO : Int := 0;   // Step number
      S_MORE : Bool := false;   // More steps are available and can be shown in S_NO
      S_ACTIVE : Bool := false;   // Step indicated in S_NO is active
      ERR_FLT : Bool := false;   // Interlock or supervision group error
      AUTO_ON : Bool := false;   // Automatic mode is active
      TAP_ON : Bool := false;   // Semiautomatic mode/step with transition enabled
      TOP_ON : Bool := false;   // Semiautomatic mode/ignore transition enabled
      MAN_ON : Bool := false;   // Manual mode is active
   END_VAR
   VAR
      HMI_INFO : Array[0..8] of UInt;
      IF_PAR : G7_IfParPlus_V6;
      RT_DATA : G7_RTDataPlus_V6;   // Internal data area
      Trans1 : G7_TransitionPlus_V6;   // Transition structure
      Trans2 : G7_TransitionPlus_V6;   // Transition structure
      Trans3 : G7_TransitionPlus_V6;   // Transition structure
      Trans4 : G7_TransitionPlus_V6;   // Transition structure
      Trans5 : G7_TransitionPlus_V6;   // Transition structure
      Trans6 : G7_TransitionPlus_V6;   // Transition structure
      Trans7 : G7_TransitionPlus_V6;   // Transition structure
      Trans8 : G7_TransitionPlus_V6;   // Transition structure
      Trans9 : G7_TransitionPlus_V6;   // Transition structure
      Trans10 : G7_TransitionPlus_V6;   // Transition structure
      Trans11 : G7_TransitionPlus_V6;   // Transition structure
      Trans12 : G7_TransitionPlus_V6;   // Transition structure
      Trans13 : G7_TransitionPlus_V6;   // Transition structure
      Trans14 : G7_TransitionPlus_V6;   // Transition structure
      "รอรับคำสั่งยา" : G7_StepPlus_V6;   // Step structure
      "Conveyorลำเลียงกล่องยาไปตำแหน่งหยิบยา" : G7_StepPlus_V6;   // Step structure
      "หมุนไปจุดเริ่มต้น" : G7_StepPlus_V6;   // Step structure
      "gripper สไลด์ออกรับยา" : G7_StepPlus_V6;   // Step structure
      "gripper หนีบกล่องยา" : G7_StepPlus_V6;   // Step structure
      "gripper สไลด์เข้า" : G7_StepPlus_V6;   // Step structure
      "gripper หมุนไปจุดปล่อย" : G7_StepPlus_V6;   // Step structure
      "แกนY เลื่อนขึ้นไปแถวที่เก็บ" : G7_StepPlus_V6;   // Step structure
      "แกนX เลื่อนไปคอลัมน์ที่เก็บ" : G7_StepPlus_V6;   // Step structure
      "gripper สไลด์ออกเพื่อปล่อยวางยา" : G7_StepPlus_V6;   // Step structure
      "gripper ปล่อยกล่องยา" : G7_StepPlus_V6;   // Step structure
      "gripper สไลด์เข้าหลังปล่อยกล่องยา" : G7_StepPlus_V6;   // Step structure
      "แกน Y เลื่อนกลับจุดเริ่มต้น" : G7_StepPlus_V6;   // Step structure
      "แกน X เลื่อนกลับจุดเริ่มต้น" : G7_StepPlus_V6;   // Step structure
      SINI : Array[0..1] of USInt;
      LSTT : Array[0..13] of USInt;
      ATAJ : Array[0..13] of USInt;
      ATAB : Array[0..13] of USInt;
      PSTT : Array[0..13] of USInt;
      NSTT : Array[0..13] of USInt;
      ASSJ : Array[0..13] of USInt;
      ASSB : Array[0..13] of USInt;
      PTTS : Array[0..13] of USInt;
      NTTS : Array[0..13] of USInt;
      SW_SQTS : Array[0..13] of USInt;
      SWITCH : Array[0..0] of USInt;
      TVX : Array[0..1] of USInt;
      TTX : Array[0..1] of USInt;
      TSX : Array[0..1] of USInt;
      S00X : Array[0..1] of USInt;
      SOFFX : Array[0..1] of USInt;
      SONX : Array[0..1] of USInt;
      SAX : Array[0..1] of USInt;
      SERRX : Array[0..14] of USInt;
      SMX : Array[0..14] of USInt;
      S0X : Array[0..14] of USInt;
      S1X : Array[0..14] of USInt;
      IL_ALARM_INST : Diag_Alarm;
      SUP_ALARM_INST : Diag_Alarm;
      STEP_TIME_ALARM_INST : Diag_Alarm;
      IEC_TIMER_INST : IEC_TIMER;
      TRANSACTION_FLAG : Bool := false;
   END_VAR
   // SINI[0] := 2;
   // LSTT[0] := 255;
   // LSTT[1] := 255;
   // LSTT[2] := 255;
   // LSTT[3] := 255;
   // LSTT[4] := 255;
   // LSTT[5] := 255;
   // LSTT[6] := 255;
   // LSTT[7] := 255;
   // LSTT[8] := 255;
   // LSTT[9] := 255;
   // LSTT[10] := 255;
   // LSTT[11] := 255;
   // LSTT[12] := 255;
   // ATAJ[1] := 1;
   // ATAJ[2] := 2;
   // ATAJ[3] := 3;
   // ATAJ[4] := 4;
   // ATAJ[5] := 5;
   // ATAJ[6] := 6;
   // ATAJ[7] := 7;
   // ATAJ[8] := 8;
   // ATAJ[9] := 9;
   // ATAJ[10] := 10;
   // ATAJ[11] := 11;
   // ATAJ[12] := 12;
   // ATAJ[13] := 13;
   // ATAB[1] := 1;
   // ATAB[2] := 2;
   // ATAB[3] := 3;
   // ATAB[4] := 4;
   // ATAB[5] := 5;
   // ATAB[6] := 6;
   // ATAB[7] := 7;
   // ATAB[8] := 8;
   // ATAB[9] := 9;
   // ATAB[10] := 10;
   // ATAB[11] := 11;
   // ATAB[12] := 12;
   // ATAB[13] := 13;
   // PSTT[1] := 1;
   // PSTT[2] := 2;
   // PSTT[3] := 3;
   // PSTT[4] := 4;
   // PSTT[5] := 5;
   // PSTT[6] := 6;
   // PSTT[7] := 7;
   // PSTT[8] := 8;
   // PSTT[9] := 9;
   // PSTT[10] := 10;
   // PSTT[11] := 11;
   // PSTT[12] := 12;
   // PSTT[13] := 13;
   // NSTT[0] := 1;
   // NSTT[1] := 2;
   // NSTT[2] := 3;
   // NSTT[3] := 4;
   // NSTT[4] := 5;
   // NSTT[5] := 6;
   // NSTT[6] := 7;
   // NSTT[7] := 8;
   // NSTT[8] := 9;
   // NSTT[9] := 10;
   // NSTT[10] := 11;
   // NSTT[11] := 12;
   // NSTT[12] := 13;
   // ASSJ[1] := 1;
   // ASSJ[2] := 2;
   // ASSJ[3] := 3;
   // ASSJ[4] := 4;
   // ASSJ[5] := 5;
   // ASSJ[6] := 6;
   // ASSJ[7] := 7;
   // ASSJ[8] := 8;
   // ASSJ[9] := 9;
   // ASSJ[10] := 10;
   // ASSJ[11] := 11;
   // ASSJ[12] := 12;
   // ASSJ[13] := 13;
   // ASSB[1] := 1;
   // ASSB[2] := 2;
   // ASSB[3] := 3;
   // ASSB[4] := 4;
   // ASSB[5] := 5;
   // ASSB[6] := 6;
   // ASSB[7] := 7;
   // ASSB[8] := 8;
   // ASSB[9] := 9;
   // ASSB[10] := 10;
   // ASSB[11] := 11;
   // ASSB[12] := 12;
   // ASSB[13] := 13;
   // PTTS[0] := 255;
   // PTTS[2] := 1;
   // PTTS[3] := 2;
   // PTTS[4] := 3;
   // PTTS[5] := 4;
   // PTTS[6] := 5;
   // PTTS[7] := 6;
   // PTTS[8] := 7;
   // PTTS[9] := 8;
   // PTTS[10] := 9;
   // PTTS[11] := 10;
   // PTTS[12] := 11;
   // PTTS[13] := 12;
   // NTTS[1] := 1;
   // NTTS[2] := 2;
   // NTTS[3] := 3;
   // NTTS[4] := 4;
   // NTTS[5] := 5;
   // NTTS[6] := 6;
   // NTTS[7] := 7;
   // NTTS[8] := 8;
   // NTTS[9] := 9;
   // NTTS[10] := 10;
   // NTTS[11] := 11;
   // NTTS[12] := 12;
   // NTTS[13] := 13;
   // TVX[0] := 16#1;
   // TTX[0] := 16#1;
   // TSX[0] := 16#1;
   // S00X[0] := 16#1;
   // SOFFX[0] := 16#1;
   // SONX[0] := 16#1;
   // SAX[0] := 16#1;
   // SERRX[0] := 16#1;
   // SMX[0] := 16#1;
   // S0X[0] := 16#1;
   // S1X[0] := 16#1;
BEGIN
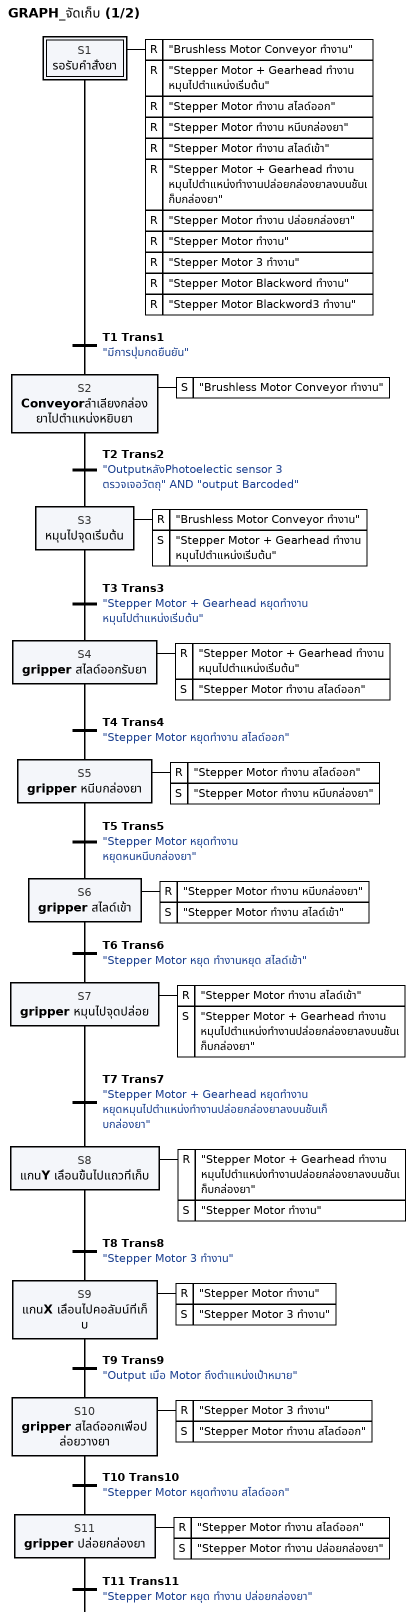
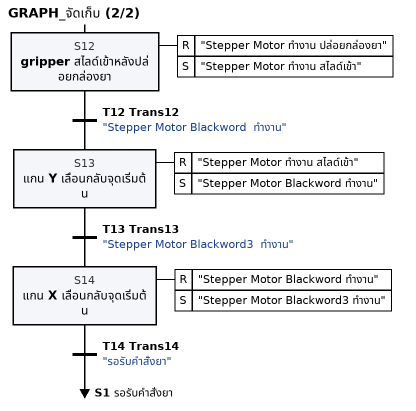
   // sequencer 1
   INITIAL_STEP "รอรับคำสั่งยา":   // S1, max time T#10S, warning time T#7S
              R    "Brushless Motor Conveyor ทำงาน"
              R    "Stepper Motor + Gearhead ทำงาน หมุนไปตำแหน่งเริ่มต้น"
              R    "Stepper Motor ทำงาน สไลด์ออก"
              R    "Stepper Motor ทำงาน หนีบกล่องยา"
              R    "Stepper Motor ทำงาน สไลด์เข้า"
              R    "Stepper Motor + Gearhead ทำงาน หมุนไปตำแหน่งทำงานปล่อยกล่องยาลงบนชั้นเก็บกล่องยา"
              R    "Stepper Motor ทำงาน ปล่อยกล่องยา"
              R    "Stepper Motor  ทำงาน"
              R    "Stepper Motor 3 ทำงาน"
              R    "Stepper Motor Blackword  ทำงาน"
              R    "Stepper Motor Blackword3  ทำงาน"
   END_STEP
   TRANSITION Trans1 FROM "รอรับคำสั่งยา" TO "Conveyorลำเลียงกล่องยาไปตำแหน่งหยิบยา"   // T1
      := "มีการปุ่มกดยืนยัน";
   END_TRANSITION
   STEP "Conveyorลำเลียงกล่องยาไปตำแหน่งหยิบยา":   // S2, max time T#10S, warning time T#7S
              S    "Brushless Motor Conveyor ทำงาน"
   END_STEP
   TRANSITION Trans2 FROM "Conveyorลำเลียงกล่องยาไปตำแหน่งหยิบยา" TO "หมุนไปจุดเริ่มต้น"   // T2
      := "OutputหลังPhotoelectic sensor 3 ตรวจเจอวัตถุ" AND "output Barcoded";
   END_TRANSITION
   STEP "หมุนไปจุดเริ่มต้น":   // S3, max time T#10S, warning time T#7S
              R    "Brushless Motor Conveyor ทำงาน"
              S    "Stepper Motor + Gearhead ทำงาน หมุนไปตำแหน่งเริ่มต้น"
   END_STEP
   TRANSITION Trans3 FROM "หมุนไปจุดเริ่มต้น" TO "gripper สไลด์ออกรับยา"   // T3
      := "Stepper Motor + Gearhead หยุดทำงาน หมุนไปตำแหน่งเริ่มต้น";
   END_TRANSITION
   STEP "gripper สไลด์ออกรับยา":   // S4, max time T#10S, warning time T#7S
              R    "Stepper Motor + Gearhead ทำงาน หมุนไปตำแหน่งเริ่มต้น"
              S    "Stepper Motor ทำงาน สไลด์ออก"
   END_STEP
   TRANSITION Trans4 FROM "gripper สไลด์ออกรับยา" TO "gripper หนีบกล่องยา"   // T4
      := "Stepper Motor หยุดทำงาน สไลด์ออก";
   END_TRANSITION
   STEP "gripper หนีบกล่องยา":   // S5, max time T#10S, warning time T#7S
              R    "Stepper Motor ทำงาน สไลด์ออก"
              S    "Stepper Motor ทำงาน หนีบกล่องยา"
   END_STEP
   TRANSITION Trans5 FROM "gripper หนีบกล่องยา" TO "gripper สไลด์เข้า"   // T5
      := "Stepper Motor หยุดทำงาน หยุดหนหนีบกล่องยา";
   END_TRANSITION
   STEP "gripper สไลด์เข้า":   // S6, max time T#10S, warning time T#7S
              R    "Stepper Motor ทำงาน หนีบกล่องยา"
              S    "Stepper Motor ทำงาน สไลด์เข้า"
   END_STEP
   TRANSITION Trans6 FROM "gripper สไลด์เข้า" TO "gripper หมุนไปจุดปล่อย"   // T6
      := "Stepper Motor หยุด ทำงานหยุด สไลด์เข้า";
   END_TRANSITION
   STEP "gripper หมุนไปจุดปล่อย":   // S7, max time T#10S, warning time T#7S
              R    "Stepper Motor ทำงาน สไลด์เข้า"
              S    "Stepper Motor + Gearhead ทำงาน หมุนไปตำแหน่งทำงานปล่อยกล่องยาลงบนชั้นเก็บกล่องยา"
   END_STEP
   TRANSITION Trans7 FROM "gripper หมุนไปจุดปล่อย" TO "แกนY เลื่อนขึ้นไปแถวที่เก็บ"   // T7
      := "Stepper Motor + Gearhead หยุดทำงาน หยุดหมุนไปตำแหน่งทำงานปล่อยกล่องยาลงบนชั้นเก็บกล่องยา";
   END_TRANSITION
   STEP "แกนY เลื่อนขึ้นไปแถวที่เก็บ":   // S8, max time T#10S, warning time T#7S
              R    "Stepper Motor + Gearhead ทำงาน หมุนไปตำแหน่งทำงานปล่อยกล่องยาลงบนชั้นเก็บกล่องยา"
              S    "Stepper Motor  ทำงาน"
   END_STEP
   TRANSITION Trans8 FROM "แกนY เลื่อนขึ้นไปแถวที่เก็บ" TO "แกนX เลื่อนไปคอลัมน์ที่เก็บ"   // T8
      := "Stepper Motor 3 ทำงาน";
   END_TRANSITION
   STEP "แกนX เลื่อนไปคอลัมน์ที่เก็บ":   // S9, max time T#10S, warning time T#7S
              R    "Stepper Motor  ทำงาน"
              S    "Stepper Motor 3 ทำงาน"
   END_STEP
   TRANSITION Trans9 FROM "แกนX เลื่อนไปคอลัมน์ที่เก็บ" TO "gripper สไลด์ออกเพื่อปล่อยวางยา"   // T9
      := "Output เมื่อ Motor ถึงตำแหน่งเป้าหมาย";
   END_TRANSITION
   STEP "gripper สไลด์ออกเพื่อปล่อยวางยา":   // S10, max time T#10S, warning time T#7S
              R    "Stepper Motor 3 ทำงาน"
              S    "Stepper Motor ทำงาน สไลด์ออก"
   END_STEP
   TRANSITION Trans10 FROM "gripper สไลด์ออกเพื่อปล่อยวางยา" TO "gripper ปล่อยกล่องยา"   // T10
      := "Stepper Motor หยุดทำงาน สไลด์ออก";
   END_TRANSITION
   STEP "gripper ปล่อยกล่องยา":   // S11, max time T#10S, warning time T#7S
              R    "Stepper Motor ทำงาน สไลด์ออก"
              S    "Stepper Motor ทำงาน ปล่อยกล่องยา"
   END_STEP
   TRANSITION Trans11 FROM "gripper ปล่อยกล่องยา" TO "gripper สไลด์เข้าหลังปล่อยกล่องยา"   // T11
      := "Stepper Motor หยุด ทำงาน ปล่อยกล่องยา";
   END_TRANSITION
   STEP "gripper สไลด์เข้าหลังปล่อยกล่องยา":   // S12, max time T#10S, warning time T#7S
              R    "Stepper Motor ทำงาน ปล่อยกล่องยา"
              S    "Stepper Motor ทำงาน สไลด์เข้า"
   END_STEP
   TRANSITION Trans12 FROM "gripper สไลด์เข้าหลังปล่อยกล่องยา" TO "แกน Y เลื่อนกลับจุดเริ่มต้น"   // T12
      := "Stepper Motor Blackword  ทำงาน";
   END_TRANSITION
   STEP "แกน Y เลื่อนกลับจุดเริ่มต้น":   // S13, max time T#10S, warning time T#7S
              R    "Stepper Motor ทำงาน สไลด์เข้า"
              S    "Stepper Motor Blackword  ทำงาน"
   END_STEP
   TRANSITION Trans13 FROM "แกน Y เลื่อนกลับจุดเริ่มต้น" TO "แกน X เลื่อนกลับจุดเริ่มต้น"   // T13
      := "Stepper Motor Blackword3  ทำงาน";
   END_TRANSITION
   STEP "แกน X เลื่อนกลับจุดเริ่มต้น":   // S14, max time T#10S, warning time T#7S
              R    "Stepper Motor Blackword  ทำงาน"
              S    "Stepper Motor Blackword3  ทำงาน"
   END_STEP
   TRANSITION Trans14 FROM "แกน X เลื่อนกลับจุดเริ่มต้น" TO "รอรับคำสั่งยา"   // T14, jump
      := "รอรับคำสั่งยา";
   END_TRANSITION
END_FUNCTION_BLOCK

FUNCTION_BLOCK "GRAPH_เบิกจ่าย"   // FB18, GRAPH_PLUS
{ S7_Optimized_Access := 'TRUE' }
VERSION : 0.1
   VAR_INPUT
      OFF_SQ : Bool := false;   // Turn sequence off
      INIT_SQ : Bool := false;   // Set sequence to initial state
      ACK_EF : Bool := false;   // Acknowledge all errors and faults
      S_PREV : Bool := false;   // Output previous step in parameter S_NO
      S_NEXT : Bool := false;   // Indicate next step in parameter S_NO
      SW_AUTO : Bool := false;   // Automatic mode
      SW_TAP : Bool := false;   // Semiautomatic/switch with transition
      SW_TOP : Bool := false;   // Semiautomatic/ignore transition
      SW_MAN : Bool := false;   // Manual mode
      S_SEL : Int := 0;   // Select step to be output to S_NO
      S_ON : Bool := false;   // Activate step indicated in S_NO
      S_OFF : Bool := false;   // Deactivate step indicated S_NO
      T_PUSH : Bool := false;   // Enable transition to switch in semi automatic mode
   END_VAR
   VAR_OUTPUT
      S_NO : Int := 0;   // Step number
      S_MORE : Bool := false;   // More steps are available and can be shown in S_NO
      S_ACTIVE : Bool := false;   // Step indicated in S_NO is active
      ERR_FLT : Bool := false;   // Interlock or supervision group error
      AUTO_ON : Bool := false;   // Automatic mode is active
      TAP_ON : Bool := false;   // Semiautomatic mode/step with transition enabled
      TOP_ON : Bool := false;   // Semiautomatic mode/ignore transition enabled
      MAN_ON : Bool := false;   // Manual mode is active
   END_VAR
   VAR
      HMI_INFO : Array[0..8] of UInt;
      IF_PAR : G7_IfParPlus_V6;
      RT_DATA : G7_RTDataPlus_V6;   // Internal data area
      Trans1 : G7_TransitionPlus_V6;   // Transition structure
      Trans2 : G7_TransitionPlus_V6;   // Transition structure
      Trans3 : G7_TransitionPlus_V6;   // Transition structure
      Trans4 : G7_TransitionPlus_V6;   // Transition structure
      Trans5 : G7_TransitionPlus_V6;   // Transition structure
      Trans6 : G7_TransitionPlus_V6;   // Transition structure
      Trans7 : G7_TransitionPlus_V6;   // Transition structure
      Trans8 : G7_TransitionPlus_V6;   // Transition structure
      "รอคำสั่งเบิกยา" : G7_StepPlus_V6;   // Step structure
      "แกน Y เลื่อนไปแถวของยา" : G7_StepPlus_V6;   // Step structure
      "แกนX เลื่อนไปคอลัมน์ของยา" : G7_StepPlus_V6;   // Step structure
      "สไลด์ตัวงัดกล่องยาออก" : G7_StepPlus_V6;   // Step structure
      "สไลด์ตัวงัดกล่องยาเข้า" : G7_StepPlus_V6;   // Step structure
      "แกน Y เลื่อนกลับจุดเริ่มต้น" : G7_StepPlus_V6;   // Step structure
      "แกนX_เลื่อนกลับจุดเริ่มต้น" : G7_StepPlus_V6;   // Step structure
      "Conveyor ลำเลียงยาไปช่องเบิกจ่าย" : G7_StepPlus_V6;   // Step structure
      SINI : Array[0..1] of USInt;
      LSTT : Array[0..7] of USInt;
      ATAJ : Array[0..7] of USInt;
      ATAB : Array[0..7] of USInt;
      PSTT : Array[0..7] of USInt;
      NSTT : Array[0..7] of USInt;
      ASSJ : Array[0..7] of USInt;
      ASSB : Array[0..7] of USInt;
      PTTS : Array[0..7] of USInt;
      NTTS : Array[0..7] of USInt;
      SW_SQTS : Array[0..7] of USInt;
      SWITCH : Array[0..0] of USInt;
      TVX : Array[0..1] of USInt;
      TTX : Array[0..1] of USInt;
      TSX : Array[0..1] of USInt;
      S00X : Array[0..1] of USInt;
      SOFFX : Array[0..1] of USInt;
      SONX : Array[0..1] of USInt;
      SAX : Array[0..1] of USInt;
      SERRX : Array[0..8] of USInt;
      SMX : Array[0..8] of USInt;
      S0X : Array[0..8] of USInt;
      S1X : Array[0..8] of USInt;
      IL_ALARM_INST : Diag_Alarm;
      SUP_ALARM_INST : Diag_Alarm;
      STEP_TIME_ALARM_INST : Diag_Alarm;
      IEC_TIMER_INST : IEC_TIMER;
      TRANSACTION_FLAG : Bool := false;
   END_VAR
   // SINI[0] := 2;
   // LSTT[0] := 255;
   // LSTT[1] := 255;
   // LSTT[2] := 255;
   // LSTT[3] := 255;
   // LSTT[4] := 255;
   // LSTT[5] := 255;
   // LSTT[6] := 255;
   // ATAJ[1] := 1;
   // ATAJ[2] := 2;
   // ATAJ[3] := 3;
   // ATAJ[4] := 4;
   // ATAJ[5] := 5;
   // ATAJ[6] := 6;
   // ATAJ[7] := 7;
   // ATAB[1] := 1;
   // ATAB[2] := 2;
   // ATAB[3] := 3;
   // ATAB[4] := 4;
   // ATAB[5] := 5;
   // ATAB[6] := 6;
   // ATAB[7] := 7;
   // PSTT[1] := 1;
   // PSTT[2] := 2;
   // PSTT[3] := 3;
   // PSTT[4] := 4;
   // PSTT[5] := 5;
   // PSTT[6] := 6;
   // PSTT[7] := 7;
   // NSTT[0] := 1;
   // NSTT[1] := 2;
   // NSTT[2] := 3;
   // NSTT[3] := 4;
   // NSTT[4] := 5;
   // NSTT[5] := 6;
   // NSTT[6] := 7;
   // ASSJ[1] := 1;
   // ASSJ[2] := 2;
   // ASSJ[3] := 3;
   // ASSJ[4] := 4;
   // ASSJ[5] := 5;
   // ASSJ[6] := 6;
   // ASSJ[7] := 7;
   // ASSB[1] := 1;
   // ASSB[2] := 2;
   // ASSB[3] := 3;
   // ASSB[4] := 4;
   // ASSB[5] := 5;
   // ASSB[6] := 6;
   // ASSB[7] := 7;
   // PTTS[0] := 255;
   // PTTS[2] := 1;
   // PTTS[3] := 2;
   // PTTS[4] := 3;
   // PTTS[5] := 4;
   // PTTS[6] := 5;
   // PTTS[7] := 6;
   // NTTS[1] := 1;
   // NTTS[2] := 2;
   // NTTS[3] := 3;
   // NTTS[4] := 4;
   // NTTS[5] := 5;
   // NTTS[6] := 6;
   // NTTS[7] := 7;
   // TVX[0] := 16#1;
   // TTX[0] := 16#1;
   // TSX[0] := 16#1;
   // S00X[0] := 16#1;
   // SOFFX[0] := 16#1;
   // SONX[0] := 16#1;
   // SAX[0] := 16#1;
   // SERRX[0] := 16#1;
   // SMX[0] := 16#1;
   // S0X[0] := 16#1;
   // S1X[0] := 16#1;
BEGIN
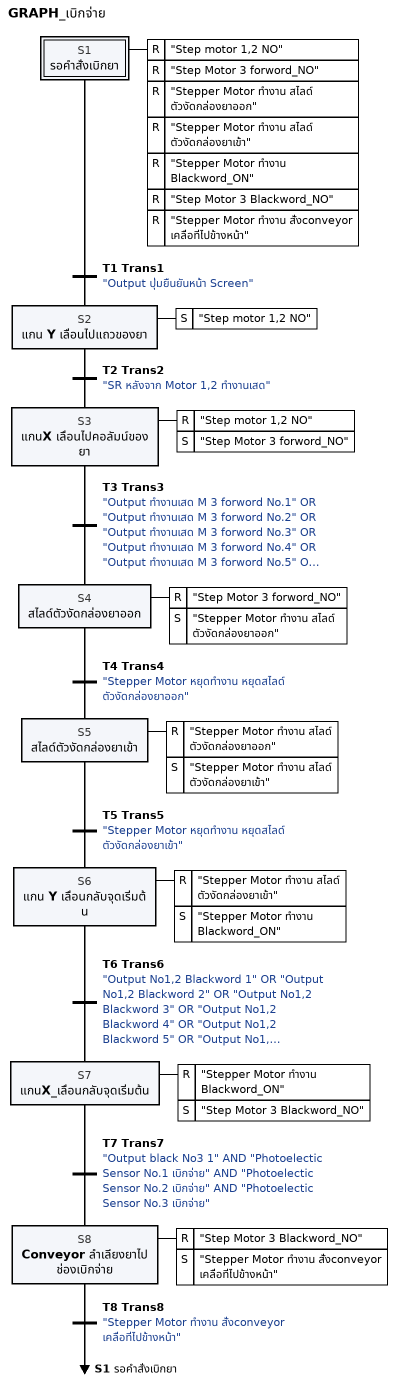
   // sequencer 1
   INITIAL_STEP "รอคำสั่งเบิกยา":   // S1, max time T#10S, warning time T#7S
              R    "Step motor 1,2 NO"
              R    "Step Motor 3 forword_NO"
              R    "Stepper Motor ทำงาน สไลด์ ตัวงัดกล่องยาออก"
              R    "Stepper Motor ทำงาน สไลด์ ตัวงัดกล่องยาเข้า"
              R    "Stepper Motor  ทำงาน Blackword_ON"
              R    "Step Motor 3 Blackword_NO"
              R    "Stepper Motor ทำงาน สั่งconveyor เคลื่อที่ไปข้างหน้า"
   END_STEP
   TRANSITION Trans1 FROM "รอคำสั่งเบิกยา" TO "แกน Y เลื่อนไปแถวของยา"   // T1
      := "Output ปุ่มยืนยันหน้า Screen";
   END_TRANSITION
   STEP "แกน Y เลื่อนไปแถวของยา":   // S2, max time T#10S, warning time T#7S
              S    "Step motor 1,2 NO"
   END_STEP
   TRANSITION Trans2 FROM "แกน Y เลื่อนไปแถวของยา" TO "แกนX เลื่อนไปคอลัมน์ของยา"   // T2
      := "SR หลังจาก Motor 1,2 ทำงานเสด";
   END_TRANSITION
   STEP "แกนX เลื่อนไปคอลัมน์ของยา":   // S3, max time T#10S, warning time T#7S
              R    "Step motor 1,2 NO"
              S    "Step Motor 3 forword_NO"
   END_STEP
   TRANSITION Trans3 FROM "แกนX เลื่อนไปคอลัมน์ของยา" TO "สไลด์ตัวงัดกล่องยาออก"   // T3
      := "Output ทำงานเสด M 3 forword No.1" OR "Output ทำงานเสด M 3 forword No.2" OR "Output ทำงานเสด M 3 forword No.3" OR "Output ทำงานเสด M 3 forword No.4" OR "Output ทำงานเสด M 3 forword No.5" OR "Output ทำงานเสด M 3 forword No.6" OR "Output ทำงานเสด M 3 forword No.7" OR "Output ทำงานเสด M 3 forword No.8" OR "Output ทำงานเสด M 3 forword No.9" OR "Output ทำงานเสด M 3 forword No.10" OR "Output ทำงานเสด M 3 forword No.11" OR "Output ทำงานเสด M 3 forword No.12" OR "Output ทำงานเสด M 3 forword No.13" OR "Output ทำงานเสด M 3 forword No.14" OR "Output ทำงานเสด M 3 forword No.15" OR "Output ทำงานเสด M 3 forword No.16" OR "Output ทำงานเสด M 3 forword No.17" OR "Output ทำงานเสด M 3 forword No.18" OR "Output ทำงานเสด M 3 forword No.19" OR "Output ทำงานเสด M 3 forword No.20" OR "Output ทำงานเสด M 3 forword No.21" OR "Output ทำงานเสด M 3 forword No.22" OR "Output ทำงานเสด M 3 forword No.23" OR "Output ทำงานเสด M 3 forword No.24" OR "Output ทำงานเสด M 3 forword No.25" OR "Output ทำงานเสด M 3 forword No.26";
   END_TRANSITION
   STEP "สไลด์ตัวงัดกล่องยาออก":   // S4, max time T#10S, warning time T#7S
              R    "Step Motor 3 forword_NO"
              S    "Stepper Motor ทำงาน สไลด์ ตัวงัดกล่องยาออก"
   END_STEP
   TRANSITION Trans4 FROM "สไลด์ตัวงัดกล่องยาออก" TO "สไลด์ตัวงัดกล่องยาเข้า"   // T4: ครบ 10 วินาที (Timer ใน FB8)
      := "Stepper Motor หยุดทำงาน หยุดสไลด์ ตัวงัดกล่องยาออก";
   END_TRANSITION
   STEP "สไลด์ตัวงัดกล่องยาเข้า":   // S5, max time T#10S, warning time T#7S
              R    "Stepper Motor ทำงาน สไลด์ ตัวงัดกล่องยาออก"
              S    "Stepper Motor ทำงาน สไลด์ ตัวงัดกล่องยาเข้า"
   END_STEP
   TRANSITION Trans5 FROM "สไลด์ตัวงัดกล่องยาเข้า" TO "แกน Y เลื่อนกลับจุดเริ่มต้น"   // T5
      := "Stepper Motor หยุดทำงาน หยุดสไลด์ ตัวงัดกล่องยาเข้า";
   END_TRANSITION
   STEP "แกน Y เลื่อนกลับจุดเริ่มต้น":   // S6, max time T#10S, warning time T#7S
              R    "Stepper Motor ทำงาน สไลด์ ตัวงัดกล่องยาเข้า"
              S    "Stepper Motor  ทำงาน Blackword_ON"
   END_STEP
   TRANSITION Trans6 FROM "แกน Y เลื่อนกลับจุดเริ่มต้น" TO "แกนX_เลื่อนกลับจุดเริ่มต้น"   // T6
      := "Output No1,2 Blackword 1" OR "Output No1,2 Blackword 2" OR "Output No1,2 Blackword 3" OR "Output No1,2 Blackword 4" OR "Output No1,2 Blackword 5" OR "Output No1,2 Blackword 6" OR "Output No1,2 Blackword 7" OR "Output No1,2 Blackword 8" OR "Output No1,2 Blackword 9" OR "Output No1,2 Blackword 10" OR "Output No1,2 Blackword 11" OR "Output No1,2 Blackword 12" OR "Output No1,2 Blackword 13" OR "Output No1,2 Blackword 14" OR "Output No1,2 Blackword 15" OR "Output No1,2 Blackword 16" OR "Output No1,2 Blackword 17" OR "Output No1,2 Blackword 18" OR "Output No1,2 Blackword 19";
   END_TRANSITION
   STEP "แกนX_เลื่อนกลับจุดเริ่มต้น":   // S7, max time T#10S, warning time T#7S
              R    "Stepper Motor  ทำงาน Blackword_ON"
              S    "Step Motor 3 Blackword_NO"
   END_STEP
   TRANSITION Trans7 FROM "แกนX_เลื่อนกลับจุดเริ่มต้น" TO "Conveyor ลำเลียงยาไปช่องเบิกจ่าย"   // T7
      := "Output black No3 1" AND "Photoelectic Sensor No.1 เบิกจ่าย" AND "Photoelectic Sensor No.2 เบิกจ่าย" AND "Photoelectic Sensor No.3 เบิกจ่าย";
   END_TRANSITION
   STEP "Conveyor ลำเลียงยาไปช่องเบิกจ่าย":   // S8, max time T#10S, warning time T#7S
              R    "Step Motor 3 Blackword_NO"
              S    "Stepper Motor ทำงาน สั่งconveyor เคลื่อที่ไปข้างหน้า"
   END_STEP
   TRANSITION Trans8 FROM "Conveyor ลำเลียงยาไปช่องเบิกจ่าย" TO "รอคำสั่งเบิกยา"   // T8, jump
      := "Stepper Motor ทำงาน สั่งconveyor เคลื่อที่ไปข้างหน้า";
   END_TRANSITION
END_FUNCTION_BLOCK

// folder: Screen หน้าจอ

FUNCTION_BLOCK "Screen Data Pro จัดเก็บ"   // FB11, LAD
{ S7_Optimized_Access := 'TRUE' }
VERSION : 0.1
   VAR_OUTPUT
      Output : Int;
   END_VAR
BEGIN

REGION Network 1
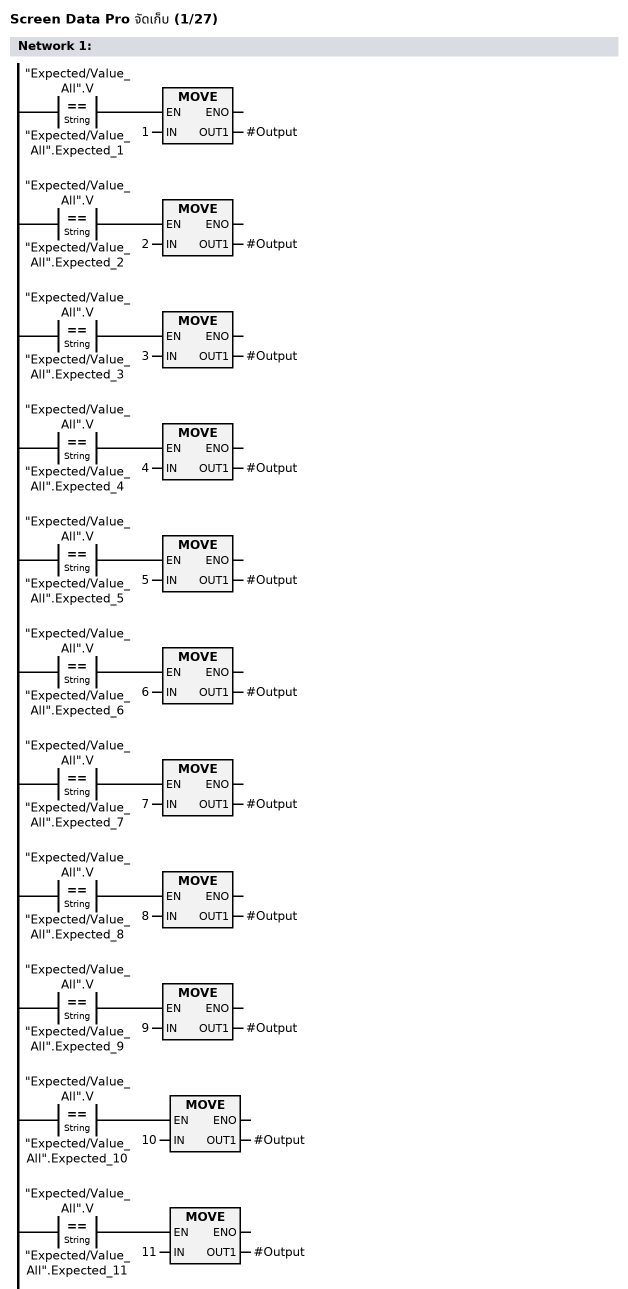
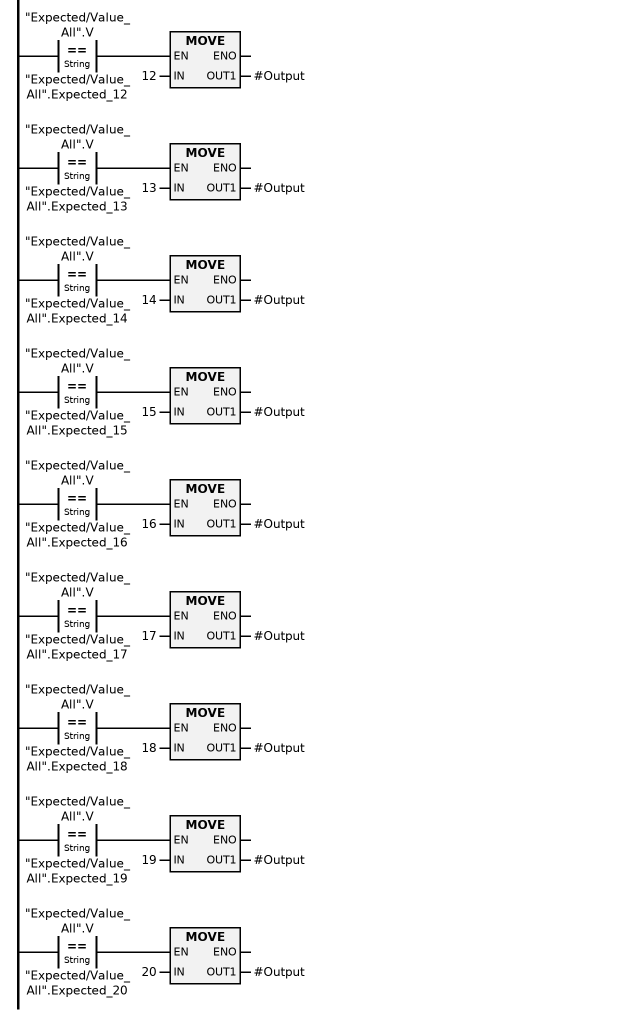
   RUNG wire#powerrail
      { S7_Templates := "SrcType := String" } EQ_Contact(in1 := "Expected/Value_All".V, in2 := "Expected/Value_All".Expected_1)
      Move(in := 1, out1 => #Output)
   END_RUNG
   RUNG wire#powerrail
      { S7_Templates := "SrcType := String" } EQ_Contact(in1 := "Expected/Value_All".V, in2 := "Expected/Value_All".Expected_2)
      Move(in := 2, out1 => #Output)
   END_RUNG
   RUNG wire#powerrail
      { S7_Templates := "SrcType := String" } EQ_Contact(in1 := "Expected/Value_All".V, in2 := "Expected/Value_All".Expected_3)
      Move(in := 3, out1 => #Output)
   END_RUNG
   RUNG wire#powerrail
      { S7_Templates := "SrcType := String" } EQ_Contact(in1 := "Expected/Value_All".V, in2 := "Expected/Value_All".Expected_4)
      Move(in := 4, out1 => #Output)
   END_RUNG
   RUNG wire#powerrail
      { S7_Templates := "SrcType := String" } EQ_Contact(in1 := "Expected/Value_All".V, in2 := "Expected/Value_All".Expected_5)
      Move(in := 5, out1 => #Output)
   END_RUNG
   RUNG wire#powerrail
      { S7_Templates := "SrcType := String" } EQ_Contact(in1 := "Expected/Value_All".V, in2 := "Expected/Value_All".Expected_6)
      Move(in := 6, out1 => #Output)
   END_RUNG
   RUNG wire#powerrail
      { S7_Templates := "SrcType := String" } EQ_Contact(in1 := "Expected/Value_All".V, in2 := "Expected/Value_All".Expected_7)
      Move(in := 7, out1 => #Output)
   END_RUNG
   RUNG wire#powerrail
      { S7_Templates := "SrcType := String" } EQ_Contact(in1 := "Expected/Value_All".V, in2 := "Expected/Value_All".Expected_8)
      Move(in := 8, out1 => #Output)
   END_RUNG
   RUNG wire#powerrail
      { S7_Templates := "SrcType := String" } EQ_Contact(in1 := "Expected/Value_All".V, in2 := "Expected/Value_All".Expected_9)
      Move(in := 9, out1 => #Output)
   END_RUNG
   RUNG wire#powerrail
      { S7_Templates := "SrcType := String" } EQ_Contact(in1 := "Expected/Value_All".V, in2 := "Expected/Value_All".Expected_10)
      Move(in := 10, out1 => #Output)
   END_RUNG
   RUNG wire#powerrail
      { S7_Templates := "SrcType := String" } EQ_Contact(in1 := "Expected/Value_All".V, in2 := "Expected/Value_All".Expected_11)
      Move(in := 11, out1 => #Output)
   END_RUNG
   RUNG wire#powerrail
      { S7_Templates := "SrcType := String" } EQ_Contact(in1 := "Expected/Value_All".V, in2 := "Expected/Value_All".Expected_12)
      Move(in := 12, out1 => #Output)
   END_RUNG
   RUNG wire#powerrail
      { S7_Templates := "SrcType := String" } EQ_Contact(in1 := "Expected/Value_All".V, in2 := "Expected/Value_All".Expected_13)
      Move(in := 13, out1 => #Output)
   END_RUNG
   RUNG wire#powerrail
      { S7_Templates := "SrcType := String" } EQ_Contact(in1 := "Expected/Value_All".V, in2 := "Expected/Value_All".Expected_14)
      Move(in := 14, out1 => #Output)
   END_RUNG
   RUNG wire#powerrail
      { S7_Templates := "SrcType := String" } EQ_Contact(in1 := "Expected/Value_All".V, in2 := "Expected/Value_All".Expected_15)
      Move(in := 15, out1 => #Output)
   END_RUNG
   RUNG wire#powerrail
      { S7_Templates := "SrcType := String" } EQ_Contact(in1 := "Expected/Value_All".V, in2 := "Expected/Value_All".Expected_16)
      Move(in := 16, out1 => #Output)
   END_RUNG
   RUNG wire#powerrail
      { S7_Templates := "SrcType := String" } EQ_Contact(in1 := "Expected/Value_All".V, in2 := "Expected/Value_All".Expected_17)
      Move(in := 17, out1 => #Output)
   END_RUNG
   RUNG wire#powerrail
      { S7_Templates := "SrcType := String" } EQ_Contact(in1 := "Expected/Value_All".V, in2 := "Expected/Value_All".Expected_18)
      Move(in := 18, out1 => #Output)
   END_RUNG
   RUNG wire#powerrail
      { S7_Templates := "SrcType := String" } EQ_Contact(in1 := "Expected/Value_All".V, in2 := "Expected/Value_All".Expected_19)
      Move(in := 19, out1 => #Output)
   END_RUNG
   RUNG wire#powerrail
      { S7_Templates := "SrcType := String" } EQ_Contact(in1 := "Expected/Value_All".V, in2 := "Expected/Value_All".Expected_20)
      Move(in := 20, out1 => #Output)
   END_RUNG
   // the same network as SCL:
   IF "Expected/Value_All".V = "Expected/Value_All".Expected_1 THEN #Output := 1; END_IF;
   IF "Expected/Value_All".V = "Expected/Value_All".Expected_2 THEN #Output := 2; END_IF;
   IF "Expected/Value_All".V = "Expected/Value_All".Expected_3 THEN #Output := 3; END_IF;
   IF "Expected/Value_All".V = "Expected/Value_All".Expected_4 THEN #Output := 4; END_IF;
   IF "Expected/Value_All".V = "Expected/Value_All".Expected_5 THEN #Output := 5; END_IF;
   IF "Expected/Value_All".V = "Expected/Value_All".Expected_6 THEN #Output := 6; END_IF;
   IF "Expected/Value_All".V = "Expected/Value_All".Expected_7 THEN #Output := 7; END_IF;
   IF "Expected/Value_All".V = "Expected/Value_All".Expected_8 THEN #Output := 8; END_IF;
   IF "Expected/Value_All".V = "Expected/Value_All".Expected_9 THEN #Output := 9; END_IF;
   IF "Expected/Value_All".V = "Expected/Value_All".Expected_10 THEN #Output := 10; END_IF;
   IF "Expected/Value_All".V = "Expected/Value_All".Expected_11 THEN #Output := 11; END_IF;
   IF "Expected/Value_All".V = "Expected/Value_All".Expected_12 THEN #Output := 12; END_IF;
   IF "Expected/Value_All".V = "Expected/Value_All".Expected_13 THEN #Output := 13; END_IF;
   IF "Expected/Value_All".V = "Expected/Value_All".Expected_14 THEN #Output := 14; END_IF;
   IF "Expected/Value_All".V = "Expected/Value_All".Expected_15 THEN #Output := 15; END_IF;
   IF "Expected/Value_All".V = "Expected/Value_All".Expected_16 THEN #Output := 16; END_IF;
   IF "Expected/Value_All".V = "Expected/Value_All".Expected_17 THEN #Output := 17; END_IF;
   IF "Expected/Value_All".V = "Expected/Value_All".Expected_18 THEN #Output := 18; END_IF;
   IF "Expected/Value_All".V = "Expected/Value_All".Expected_19 THEN #Output := 19; END_IF;
   IF "Expected/Value_All".V = "Expected/Value_All".Expected_20 THEN #Output := 20; END_IF;
END_REGION

REGION Network 2
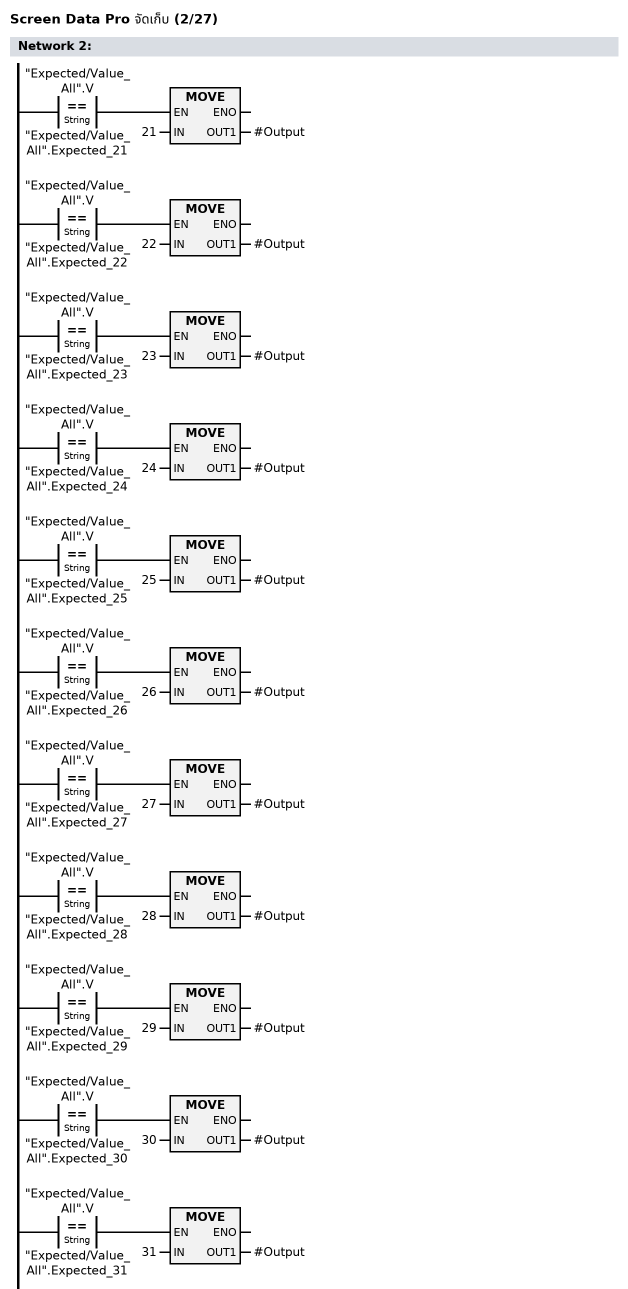
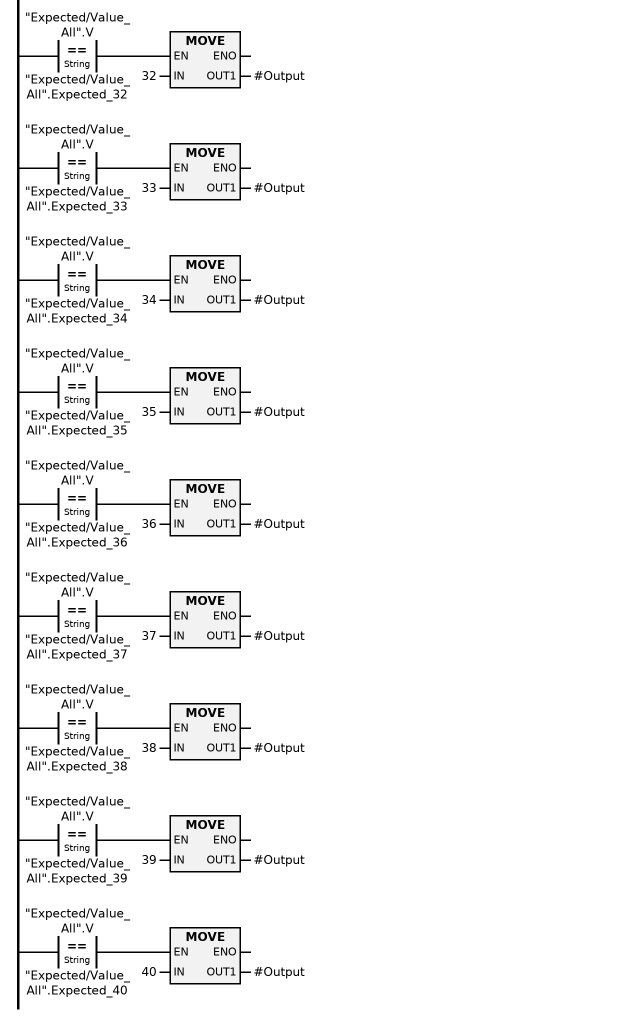
   RUNG wire#powerrail
      { S7_Templates := "SrcType := String" } EQ_Contact(in1 := "Expected/Value_All".V, in2 := "Expected/Value_All".Expected_21)
      Move(in := 21, out1 => #Output)
   END_RUNG
   RUNG wire#powerrail
      { S7_Templates := "SrcType := String" } EQ_Contact(in1 := "Expected/Value_All".V, in2 := "Expected/Value_All".Expected_22)
      Move(in := 22, out1 => #Output)
   END_RUNG
   RUNG wire#powerrail
      { S7_Templates := "SrcType := String" } EQ_Contact(in1 := "Expected/Value_All".V, in2 := "Expected/Value_All".Expected_23)
      Move(in := 23, out1 => #Output)
   END_RUNG
   RUNG wire#powerrail
      { S7_Templates := "SrcType := String" } EQ_Contact(in1 := "Expected/Value_All".V, in2 := "Expected/Value_All".Expected_24)
      Move(in := 24, out1 => #Output)
   END_RUNG
   RUNG wire#powerrail
      { S7_Templates := "SrcType := String" } EQ_Contact(in1 := "Expected/Value_All".V, in2 := "Expected/Value_All".Expected_25)
      Move(in := 25, out1 => #Output)
   END_RUNG
   RUNG wire#powerrail
      { S7_Templates := "SrcType := String" } EQ_Contact(in1 := "Expected/Value_All".V, in2 := "Expected/Value_All".Expected_26)
      Move(in := 26, out1 => #Output)
   END_RUNG
   RUNG wire#powerrail
      { S7_Templates := "SrcType := String" } EQ_Contact(in1 := "Expected/Value_All".V, in2 := "Expected/Value_All".Expected_27)
      Move(in := 27, out1 => #Output)
   END_RUNG
   RUNG wire#powerrail
      { S7_Templates := "SrcType := String" } EQ_Contact(in1 := "Expected/Value_All".V, in2 := "Expected/Value_All".Expected_28)
      Move(in := 28, out1 => #Output)
   END_RUNG
   RUNG wire#powerrail
      { S7_Templates := "SrcType := String" } EQ_Contact(in1 := "Expected/Value_All".V, in2 := "Expected/Value_All".Expected_29)
      Move(in := 29, out1 => #Output)
   END_RUNG
   RUNG wire#powerrail
      { S7_Templates := "SrcType := String" } EQ_Contact(in1 := "Expected/Value_All".V, in2 := "Expected/Value_All".Expected_30)
      Move(in := 30, out1 => #Output)
   END_RUNG
   RUNG wire#powerrail
      { S7_Templates := "SrcType := String" } EQ_Contact(in1 := "Expected/Value_All".V, in2 := "Expected/Value_All".Expected_31)
      Move(in := 31, out1 => #Output)
   END_RUNG
   RUNG wire#powerrail
      { S7_Templates := "SrcType := String" } EQ_Contact(in1 := "Expected/Value_All".V, in2 := "Expected/Value_All".Expected_32)
      Move(in := 32, out1 => #Output)
   END_RUNG
   RUNG wire#powerrail
      { S7_Templates := "SrcType := String" } EQ_Contact(in1 := "Expected/Value_All".V, in2 := "Expected/Value_All".Expected_33)
      Move(in := 33, out1 => #Output)
   END_RUNG
   RUNG wire#powerrail
      { S7_Templates := "SrcType := String" } EQ_Contact(in1 := "Expected/Value_All".V, in2 := "Expected/Value_All".Expected_34)
      Move(in := 34, out1 => #Output)
   END_RUNG
   RUNG wire#powerrail
      { S7_Templates := "SrcType := String" } EQ_Contact(in1 := "Expected/Value_All".V, in2 := "Expected/Value_All".Expected_35)
      Move(in := 35, out1 => #Output)
   END_RUNG
   RUNG wire#powerrail
      { S7_Templates := "SrcType := String" } EQ_Contact(in1 := "Expected/Value_All".V, in2 := "Expected/Value_All".Expected_36)
      Move(in := 36, out1 => #Output)
   END_RUNG
   RUNG wire#powerrail
      { S7_Templates := "SrcType := String" } EQ_Contact(in1 := "Expected/Value_All".V, in2 := "Expected/Value_All".Expected_37)
      Move(in := 37, out1 => #Output)
   END_RUNG
   RUNG wire#powerrail
      { S7_Templates := "SrcType := String" } EQ_Contact(in1 := "Expected/Value_All".V, in2 := "Expected/Value_All".Expected_38)
      Move(in := 38, out1 => #Output)
   END_RUNG
   RUNG wire#powerrail
      { S7_Templates := "SrcType := String" } EQ_Contact(in1 := "Expected/Value_All".V, in2 := "Expected/Value_All".Expected_39)
      Move(in := 39, out1 => #Output)
   END_RUNG
   RUNG wire#powerrail
      { S7_Templates := "SrcType := String" } EQ_Contact(in1 := "Expected/Value_All".V, in2 := "Expected/Value_All".Expected_40)
      Move(in := 40, out1 => #Output)
   END_RUNG
   // the same network as SCL:
   IF "Expected/Value_All".V = "Expected/Value_All".Expected_21 THEN #Output := 21; END_IF;
   IF "Expected/Value_All".V = "Expected/Value_All".Expected_22 THEN #Output := 22; END_IF;
   IF "Expected/Value_All".V = "Expected/Value_All".Expected_23 THEN #Output := 23; END_IF;
   IF "Expected/Value_All".V = "Expected/Value_All".Expected_24 THEN #Output := 24; END_IF;
   IF "Expected/Value_All".V = "Expected/Value_All".Expected_25 THEN #Output := 25; END_IF;
   IF "Expected/Value_All".V = "Expected/Value_All".Expected_26 THEN #Output := 26; END_IF;
   IF "Expected/Value_All".V = "Expected/Value_All".Expected_27 THEN #Output := 27; END_IF;
   IF "Expected/Value_All".V = "Expected/Value_All".Expected_28 THEN #Output := 28; END_IF;
   IF "Expected/Value_All".V = "Expected/Value_All".Expected_29 THEN #Output := 29; END_IF;
   IF "Expected/Value_All".V = "Expected/Value_All".Expected_30 THEN #Output := 30; END_IF;
   IF "Expected/Value_All".V = "Expected/Value_All".Expected_31 THEN #Output := 31; END_IF;
   IF "Expected/Value_All".V = "Expected/Value_All".Expected_32 THEN #Output := 32; END_IF;
   IF "Expected/Value_All".V = "Expected/Value_All".Expected_33 THEN #Output := 33; END_IF;
   IF "Expected/Value_All".V = "Expected/Value_All".Expected_34 THEN #Output := 34; END_IF;
   IF "Expected/Value_All".V = "Expected/Value_All".Expected_35 THEN #Output := 35; END_IF;
   IF "Expected/Value_All".V = "Expected/Value_All".Expected_36 THEN #Output := 36; END_IF;
   IF "Expected/Value_All".V = "Expected/Value_All".Expected_37 THEN #Output := 37; END_IF;
   IF "Expected/Value_All".V = "Expected/Value_All".Expected_38 THEN #Output := 38; END_IF;
   IF "Expected/Value_All".V = "Expected/Value_All".Expected_39 THEN #Output := 39; END_IF;
   IF "Expected/Value_All".V = "Expected/Value_All".Expected_40 THEN #Output := 40; END_IF;
END_REGION

REGION Network 3
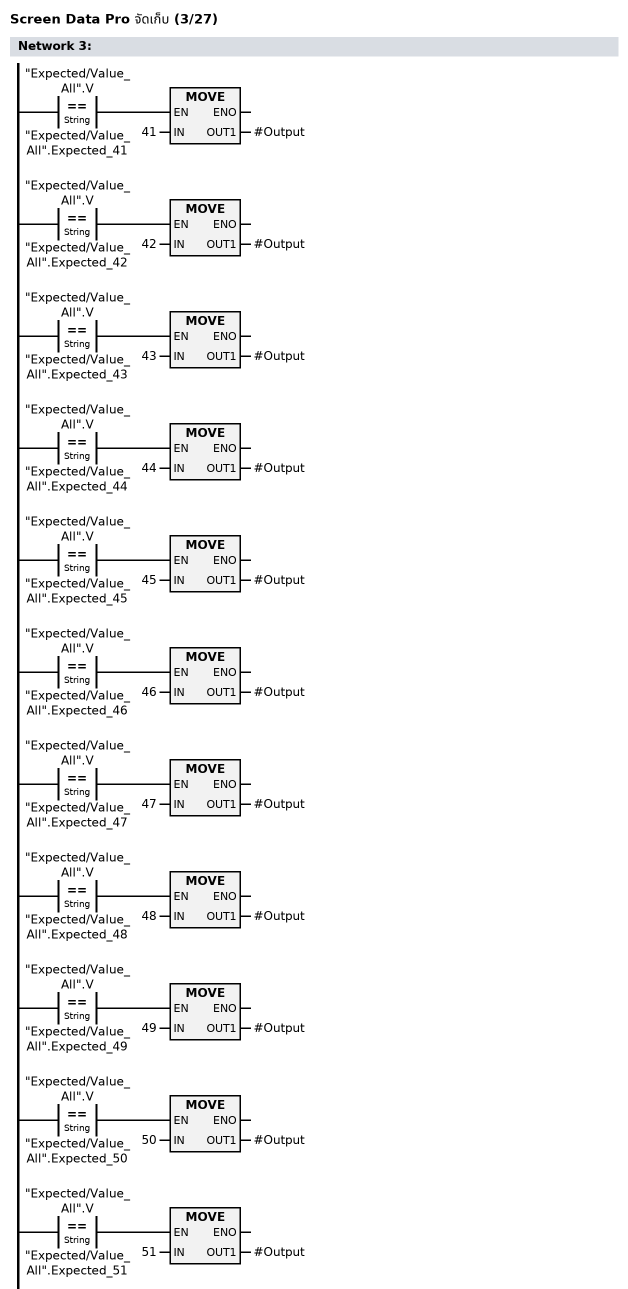
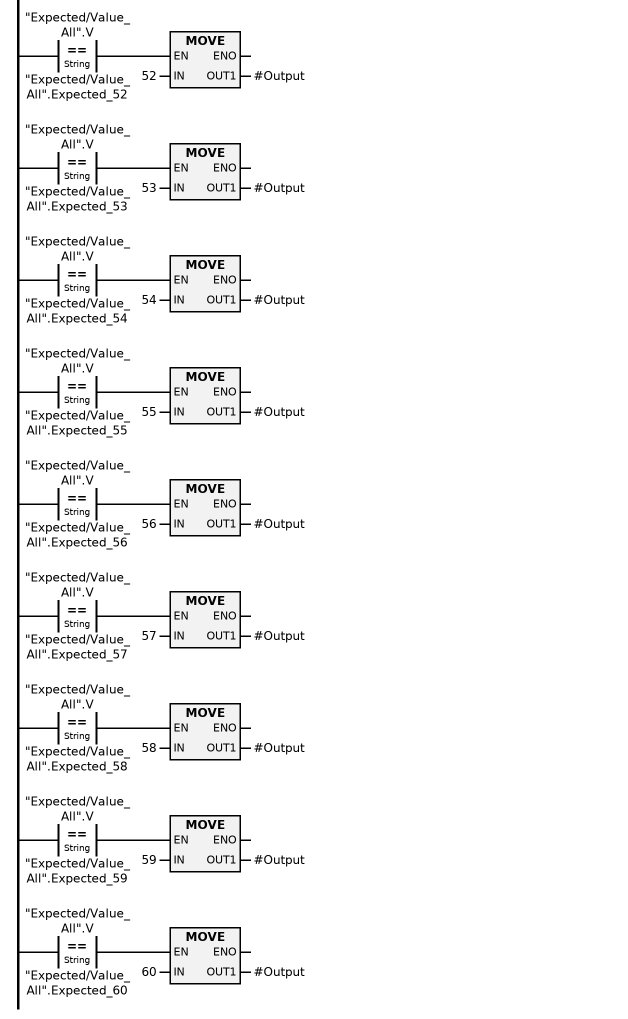
   RUNG wire#powerrail
      { S7_Templates := "SrcType := String" } EQ_Contact(in1 := "Expected/Value_All".V, in2 := "Expected/Value_All".Expected_41)
      Move(in := 41, out1 => #Output)
   END_RUNG
   RUNG wire#powerrail
      { S7_Templates := "SrcType := String" } EQ_Contact(in1 := "Expected/Value_All".V, in2 := "Expected/Value_All".Expected_42)
      Move(in := 42, out1 => #Output)
   END_RUNG
   RUNG wire#powerrail
      { S7_Templates := "SrcType := String" } EQ_Contact(in1 := "Expected/Value_All".V, in2 := "Expected/Value_All".Expected_43)
      Move(in := 43, out1 => #Output)
   END_RUNG
   RUNG wire#powerrail
      { S7_Templates := "SrcType := String" } EQ_Contact(in1 := "Expected/Value_All".V, in2 := "Expected/Value_All".Expected_44)
      Move(in := 44, out1 => #Output)
   END_RUNG
   RUNG wire#powerrail
      { S7_Templates := "SrcType := String" } EQ_Contact(in1 := "Expected/Value_All".V, in2 := "Expected/Value_All".Expected_45)
      Move(in := 45, out1 => #Output)
   END_RUNG
   RUNG wire#powerrail
      { S7_Templates := "SrcType := String" } EQ_Contact(in1 := "Expected/Value_All".V, in2 := "Expected/Value_All".Expected_46)
      Move(in := 46, out1 => #Output)
   END_RUNG
   RUNG wire#powerrail
      { S7_Templates := "SrcType := String" } EQ_Contact(in1 := "Expected/Value_All".V, in2 := "Expected/Value_All".Expected_47)
      Move(in := 47, out1 => #Output)
   END_RUNG
   RUNG wire#powerrail
      { S7_Templates := "SrcType := String" } EQ_Contact(in1 := "Expected/Value_All".V, in2 := "Expected/Value_All".Expected_48)
      Move(in := 48, out1 => #Output)
   END_RUNG
   RUNG wire#powerrail
      { S7_Templates := "SrcType := String" } EQ_Contact(in1 := "Expected/Value_All".V, in2 := "Expected/Value_All".Expected_49)
      Move(in := 49, out1 => #Output)
   END_RUNG
   RUNG wire#powerrail
      { S7_Templates := "SrcType := String" } EQ_Contact(in1 := "Expected/Value_All".V, in2 := "Expected/Value_All".Expected_50)
      Move(in := 50, out1 => #Output)
   END_RUNG
   RUNG wire#powerrail
      { S7_Templates := "SrcType := String" } EQ_Contact(in1 := "Expected/Value_All".V, in2 := "Expected/Value_All".Expected_51)
      Move(in := 51, out1 => #Output)
   END_RUNG
   RUNG wire#powerrail
      { S7_Templates := "SrcType := String" } EQ_Contact(in1 := "Expected/Value_All".V, in2 := "Expected/Value_All".Expected_52)
      Move(in := 52, out1 => #Output)
   END_RUNG
   RUNG wire#powerrail
      { S7_Templates := "SrcType := String" } EQ_Contact(in1 := "Expected/Value_All".V, in2 := "Expected/Value_All".Expected_53)
      Move(in := 53, out1 => #Output)
   END_RUNG
   RUNG wire#powerrail
      { S7_Templates := "SrcType := String" } EQ_Contact(in1 := "Expected/Value_All".V, in2 := "Expected/Value_All".Expected_54)
      Move(in := 54, out1 => #Output)
   END_RUNG
   RUNG wire#powerrail
      { S7_Templates := "SrcType := String" } EQ_Contact(in1 := "Expected/Value_All".V, in2 := "Expected/Value_All".Expected_55)
      Move(in := 55, out1 => #Output)
   END_RUNG
   RUNG wire#powerrail
      { S7_Templates := "SrcType := String" } EQ_Contact(in1 := "Expected/Value_All".V, in2 := "Expected/Value_All".Expected_56)
      Move(in := 56, out1 => #Output)
   END_RUNG
   RUNG wire#powerrail
      { S7_Templates := "SrcType := String" } EQ_Contact(in1 := "Expected/Value_All".V, in2 := "Expected/Value_All".Expected_57)
      Move(in := 57, out1 => #Output)
   END_RUNG
   RUNG wire#powerrail
      { S7_Templates := "SrcType := String" } EQ_Contact(in1 := "Expected/Value_All".V, in2 := "Expected/Value_All".Expected_58)
      Move(in := 58, out1 => #Output)
   END_RUNG
   RUNG wire#powerrail
      { S7_Templates := "SrcType := String" } EQ_Contact(in1 := "Expected/Value_All".V, in2 := "Expected/Value_All".Expected_59)
      Move(in := 59, out1 => #Output)
   END_RUNG
   RUNG wire#powerrail
      { S7_Templates := "SrcType := String" } EQ_Contact(in1 := "Expected/Value_All".V, in2 := "Expected/Value_All".Expected_60)
      Move(in := 60, out1 => #Output)
   END_RUNG
   // the same network as SCL:
   IF "Expected/Value_All".V = "Expected/Value_All".Expected_41 THEN #Output := 41; END_IF;
   IF "Expected/Value_All".V = "Expected/Value_All".Expected_42 THEN #Output := 42; END_IF;
   IF "Expected/Value_All".V = "Expected/Value_All".Expected_43 THEN #Output := 43; END_IF;
   IF "Expected/Value_All".V = "Expected/Value_All".Expected_44 THEN #Output := 44; END_IF;
   IF "Expected/Value_All".V = "Expected/Value_All".Expected_45 THEN #Output := 45; END_IF;
   IF "Expected/Value_All".V = "Expected/Value_All".Expected_46 THEN #Output := 46; END_IF;
   IF "Expected/Value_All".V = "Expected/Value_All".Expected_47 THEN #Output := 47; END_IF;
   IF "Expected/Value_All".V = "Expected/Value_All".Expected_48 THEN #Output := 48; END_IF;
   IF "Expected/Value_All".V = "Expected/Value_All".Expected_49 THEN #Output := 49; END_IF;
   IF "Expected/Value_All".V = "Expected/Value_All".Expected_50 THEN #Output := 50; END_IF;
   IF "Expected/Value_All".V = "Expected/Value_All".Expected_51 THEN #Output := 51; END_IF;
   IF "Expected/Value_All".V = "Expected/Value_All".Expected_52 THEN #Output := 52; END_IF;
   IF "Expected/Value_All".V = "Expected/Value_All".Expected_53 THEN #Output := 53; END_IF;
   IF "Expected/Value_All".V = "Expected/Value_All".Expected_54 THEN #Output := 54; END_IF;
   IF "Expected/Value_All".V = "Expected/Value_All".Expected_55 THEN #Output := 55; END_IF;
   IF "Expected/Value_All".V = "Expected/Value_All".Expected_56 THEN #Output := 56; END_IF;
   IF "Expected/Value_All".V = "Expected/Value_All".Expected_57 THEN #Output := 57; END_IF;
   IF "Expected/Value_All".V = "Expected/Value_All".Expected_58 THEN #Output := 58; END_IF;
   IF "Expected/Value_All".V = "Expected/Value_All".Expected_59 THEN #Output := 59; END_IF;
   IF "Expected/Value_All".V = "Expected/Value_All".Expected_60 THEN #Output := 60; END_IF;
END_REGION

REGION Network 4
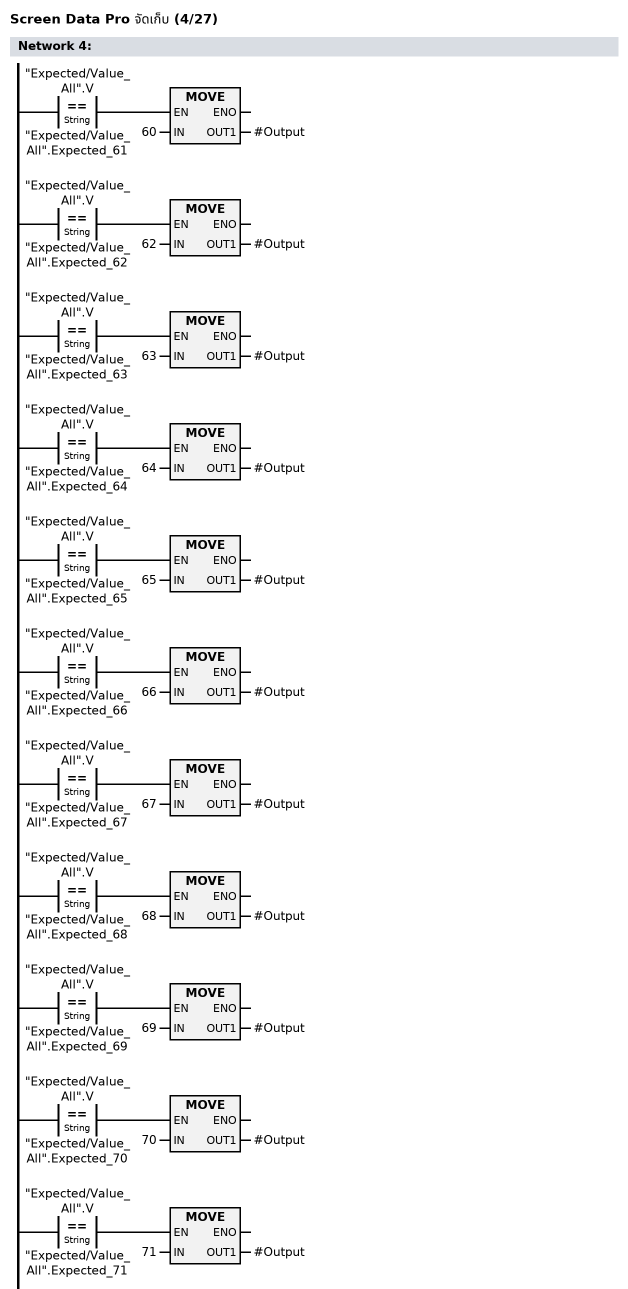
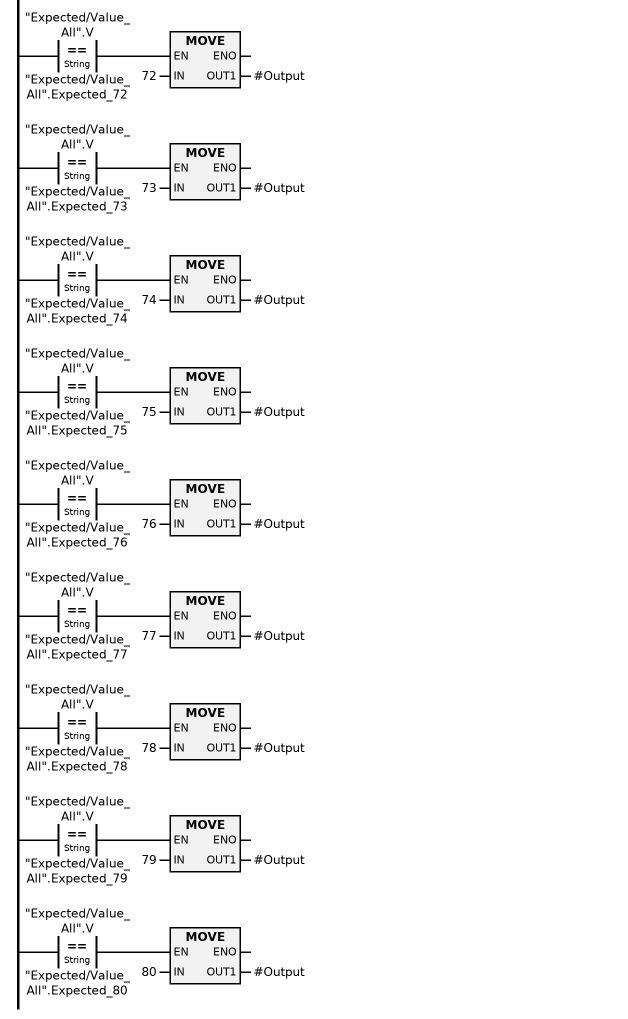
   RUNG wire#powerrail
      { S7_Templates := "SrcType := String" } EQ_Contact(in1 := "Expected/Value_All".V, in2 := "Expected/Value_All".Expected_61)
      Move(in := 60, out1 => #Output)
   END_RUNG
   RUNG wire#powerrail
      { S7_Templates := "SrcType := String" } EQ_Contact(in1 := "Expected/Value_All".V, in2 := "Expected/Value_All".Expected_62)
      Move(in := 62, out1 => #Output)
   END_RUNG
   RUNG wire#powerrail
      { S7_Templates := "SrcType := String" } EQ_Contact(in1 := "Expected/Value_All".V, in2 := "Expected/Value_All".Expected_63)
      Move(in := 63, out1 => #Output)
   END_RUNG
   RUNG wire#powerrail
      { S7_Templates := "SrcType := String" } EQ_Contact(in1 := "Expected/Value_All".V, in2 := "Expected/Value_All".Expected_64)
      Move(in := 64, out1 => #Output)
   END_RUNG
   RUNG wire#powerrail
      { S7_Templates := "SrcType := String" } EQ_Contact(in1 := "Expected/Value_All".V, in2 := "Expected/Value_All".Expected_65)
      Move(in := 65, out1 => #Output)
   END_RUNG
   RUNG wire#powerrail
      { S7_Templates := "SrcType := String" } EQ_Contact(in1 := "Expected/Value_All".V, in2 := "Expected/Value_All".Expected_66)
      Move(in := 66, out1 => #Output)
   END_RUNG
   RUNG wire#powerrail
      { S7_Templates := "SrcType := String" } EQ_Contact(in1 := "Expected/Value_All".V, in2 := "Expected/Value_All".Expected_67)
      Move(in := 67, out1 => #Output)
   END_RUNG
   RUNG wire#powerrail
      { S7_Templates := "SrcType := String" } EQ_Contact(in1 := "Expected/Value_All".V, in2 := "Expected/Value_All".Expected_68)
      Move(in := 68, out1 => #Output)
   END_RUNG
   RUNG wire#powerrail
      { S7_Templates := "SrcType := String" } EQ_Contact(in1 := "Expected/Value_All".V, in2 := "Expected/Value_All".Expected_69)
      Move(in := 69, out1 => #Output)
   END_RUNG
   RUNG wire#powerrail
      { S7_Templates := "SrcType := String" } EQ_Contact(in1 := "Expected/Value_All".V, in2 := "Expected/Value_All".Expected_70)
      Move(in := 70, out1 => #Output)
   END_RUNG
   RUNG wire#powerrail
      { S7_Templates := "SrcType := String" } EQ_Contact(in1 := "Expected/Value_All".V, in2 := "Expected/Value_All".Expected_71)
      Move(in := 71, out1 => #Output)
   END_RUNG
   RUNG wire#powerrail
      { S7_Templates := "SrcType := String" } EQ_Contact(in1 := "Expected/Value_All".V, in2 := "Expected/Value_All".Expected_72)
      Move(in := 72, out1 => #Output)
   END_RUNG
   RUNG wire#powerrail
      { S7_Templates := "SrcType := String" } EQ_Contact(in1 := "Expected/Value_All".V, in2 := "Expected/Value_All".Expected_73)
      Move(in := 73, out1 => #Output)
   END_RUNG
   RUNG wire#powerrail
      { S7_Templates := "SrcType := String" } EQ_Contact(in1 := "Expected/Value_All".V, in2 := "Expected/Value_All".Expected_74)
      Move(in := 74, out1 => #Output)
   END_RUNG
   RUNG wire#powerrail
      { S7_Templates := "SrcType := String" } EQ_Contact(in1 := "Expected/Value_All".V, in2 := "Expected/Value_All".Expected_75)
      Move(in := 75, out1 => #Output)
   END_RUNG
   RUNG wire#powerrail
      { S7_Templates := "SrcType := String" } EQ_Contact(in1 := "Expected/Value_All".V, in2 := "Expected/Value_All".Expected_76)
      Move(in := 76, out1 => #Output)
   END_RUNG
   RUNG wire#powerrail
      { S7_Templates := "SrcType := String" } EQ_Contact(in1 := "Expected/Value_All".V, in2 := "Expected/Value_All".Expected_77)
      Move(in := 77, out1 => #Output)
   END_RUNG
   RUNG wire#powerrail
      { S7_Templates := "SrcType := String" } EQ_Contact(in1 := "Expected/Value_All".V, in2 := "Expected/Value_All".Expected_78)
      Move(in := 78, out1 => #Output)
   END_RUNG
   RUNG wire#powerrail
      { S7_Templates := "SrcType := String" } EQ_Contact(in1 := "Expected/Value_All".V, in2 := "Expected/Value_All".Expected_79)
      Move(in := 79, out1 => #Output)
   END_RUNG
   RUNG wire#powerrail
      { S7_Templates := "SrcType := String" } EQ_Contact(in1 := "Expected/Value_All".V, in2 := "Expected/Value_All".Expected_80)
      Move(in := 80, out1 => #Output)
   END_RUNG
   // the same network as SCL:
   IF "Expected/Value_All".V = "Expected/Value_All".Expected_61 THEN #Output := 60; END_IF;
   IF "Expected/Value_All".V = "Expected/Value_All".Expected_62 THEN #Output := 62; END_IF;
   IF "Expected/Value_All".V = "Expected/Value_All".Expected_63 THEN #Output := 63; END_IF;
   IF "Expected/Value_All".V = "Expected/Value_All".Expected_64 THEN #Output := 64; END_IF;
   IF "Expected/Value_All".V = "Expected/Value_All".Expected_65 THEN #Output := 65; END_IF;
   IF "Expected/Value_All".V = "Expected/Value_All".Expected_66 THEN #Output := 66; END_IF;
   IF "Expected/Value_All".V = "Expected/Value_All".Expected_67 THEN #Output := 67; END_IF;
   IF "Expected/Value_All".V = "Expected/Value_All".Expected_68 THEN #Output := 68; END_IF;
   IF "Expected/Value_All".V = "Expected/Value_All".Expected_69 THEN #Output := 69; END_IF;
   IF "Expected/Value_All".V = "Expected/Value_All".Expected_70 THEN #Output := 70; END_IF;
   IF "Expected/Value_All".V = "Expected/Value_All".Expected_71 THEN #Output := 71; END_IF;
   IF "Expected/Value_All".V = "Expected/Value_All".Expected_72 THEN #Output := 72; END_IF;
   IF "Expected/Value_All".V = "Expected/Value_All".Expected_73 THEN #Output := 73; END_IF;
   IF "Expected/Value_All".V = "Expected/Value_All".Expected_74 THEN #Output := 74; END_IF;
   IF "Expected/Value_All".V = "Expected/Value_All".Expected_75 THEN #Output := 75; END_IF;
   IF "Expected/Value_All".V = "Expected/Value_All".Expected_76 THEN #Output := 76; END_IF;
   IF "Expected/Value_All".V = "Expected/Value_All".Expected_77 THEN #Output := 77; END_IF;
   IF "Expected/Value_All".V = "Expected/Value_All".Expected_78 THEN #Output := 78; END_IF;
   IF "Expected/Value_All".V = "Expected/Value_All".Expected_79 THEN #Output := 79; END_IF;
   IF "Expected/Value_All".V = "Expected/Value_All".Expected_80 THEN #Output := 80; END_IF;
END_REGION

REGION Network 5
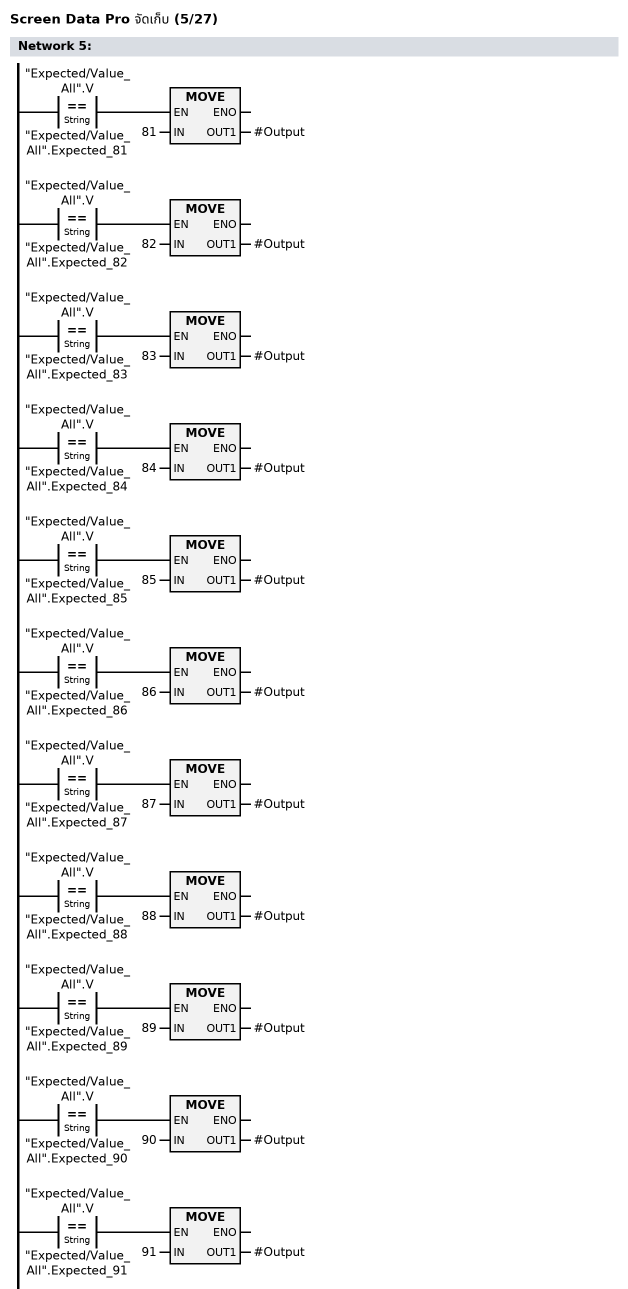
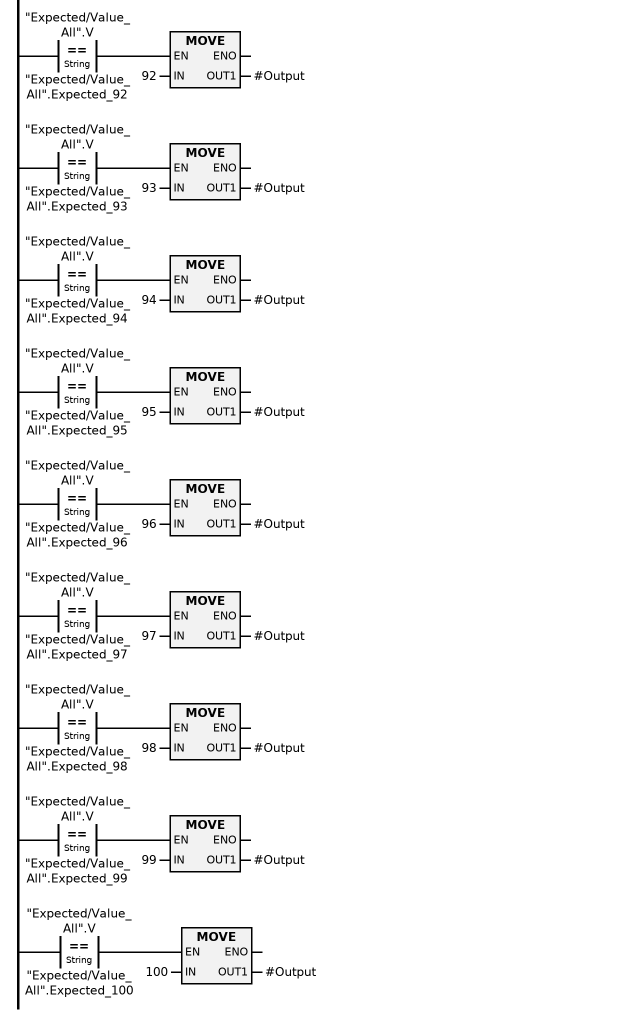
   RUNG wire#powerrail
      { S7_Templates := "SrcType := String" } EQ_Contact(in1 := "Expected/Value_All".V, in2 := "Expected/Value_All".Expected_81)
      Move(in := 81, out1 => #Output)
   END_RUNG
   RUNG wire#powerrail
      { S7_Templates := "SrcType := String" } EQ_Contact(in1 := "Expected/Value_All".V, in2 := "Expected/Value_All".Expected_82)
      Move(in := 82, out1 => #Output)
   END_RUNG
   RUNG wire#powerrail
      { S7_Templates := "SrcType := String" } EQ_Contact(in1 := "Expected/Value_All".V, in2 := "Expected/Value_All".Expected_83)
      Move(in := 83, out1 => #Output)
   END_RUNG
   RUNG wire#powerrail
      { S7_Templates := "SrcType := String" } EQ_Contact(in1 := "Expected/Value_All".V, in2 := "Expected/Value_All".Expected_84)
      Move(in := 84, out1 => #Output)
   END_RUNG
   RUNG wire#powerrail
      { S7_Templates := "SrcType := String" } EQ_Contact(in1 := "Expected/Value_All".V, in2 := "Expected/Value_All".Expected_85)
      Move(in := 85, out1 => #Output)
   END_RUNG
   RUNG wire#powerrail
      { S7_Templates := "SrcType := String" } EQ_Contact(in1 := "Expected/Value_All".V, in2 := "Expected/Value_All".Expected_86)
      Move(in := 86, out1 => #Output)
   END_RUNG
   RUNG wire#powerrail
      { S7_Templates := "SrcType := String" } EQ_Contact(in1 := "Expected/Value_All".V, in2 := "Expected/Value_All".Expected_87)
      Move(in := 87, out1 => #Output)
   END_RUNG
   RUNG wire#powerrail
      { S7_Templates := "SrcType := String" } EQ_Contact(in1 := "Expected/Value_All".V, in2 := "Expected/Value_All".Expected_88)
      Move(in := 88, out1 => #Output)
   END_RUNG
   RUNG wire#powerrail
      { S7_Templates := "SrcType := String" } EQ_Contact(in1 := "Expected/Value_All".V, in2 := "Expected/Value_All".Expected_89)
      Move(in := 89, out1 => #Output)
   END_RUNG
   RUNG wire#powerrail
      { S7_Templates := "SrcType := String" } EQ_Contact(in1 := "Expected/Value_All".V, in2 := "Expected/Value_All".Expected_90)
      Move(in := 90, out1 => #Output)
   END_RUNG
   RUNG wire#powerrail
      { S7_Templates := "SrcType := String" } EQ_Contact(in1 := "Expected/Value_All".V, in2 := "Expected/Value_All".Expected_91)
      Move(in := 91, out1 => #Output)
   END_RUNG
   RUNG wire#powerrail
      { S7_Templates := "SrcType := String" } EQ_Contact(in1 := "Expected/Value_All".V, in2 := "Expected/Value_All".Expected_92)
      Move(in := 92, out1 => #Output)
   END_RUNG
   RUNG wire#powerrail
      { S7_Templates := "SrcType := String" } EQ_Contact(in1 := "Expected/Value_All".V, in2 := "Expected/Value_All".Expected_93)
      Move(in := 93, out1 => #Output)
   END_RUNG
   RUNG wire#powerrail
      { S7_Templates := "SrcType := String" } EQ_Contact(in1 := "Expected/Value_All".V, in2 := "Expected/Value_All".Expected_94)
      Move(in := 94, out1 => #Output)
   END_RUNG
   RUNG wire#powerrail
      { S7_Templates := "SrcType := String" } EQ_Contact(in1 := "Expected/Value_All".V, in2 := "Expected/Value_All".Expected_95)
      Move(in := 95, out1 => #Output)
   END_RUNG
   RUNG wire#powerrail
      { S7_Templates := "SrcType := String" } EQ_Contact(in1 := "Expected/Value_All".V, in2 := "Expected/Value_All".Expected_96)
      Move(in := 96, out1 => #Output)
   END_RUNG
   RUNG wire#powerrail
      { S7_Templates := "SrcType := String" } EQ_Contact(in1 := "Expected/Value_All".V, in2 := "Expected/Value_All".Expected_97)
      Move(in := 97, out1 => #Output)
   END_RUNG
   RUNG wire#powerrail
      { S7_Templates := "SrcType := String" } EQ_Contact(in1 := "Expected/Value_All".V, in2 := "Expected/Value_All".Expected_98)
      Move(in := 98, out1 => #Output)
   END_RUNG
   RUNG wire#powerrail
      { S7_Templates := "SrcType := String" } EQ_Contact(in1 := "Expected/Value_All".V, in2 := "Expected/Value_All".Expected_99)
      Move(in := 99, out1 => #Output)
   END_RUNG
   RUNG wire#powerrail
      { S7_Templates := "SrcType := String" } EQ_Contact(in1 := "Expected/Value_All".V, in2 := "Expected/Value_All".Expected_100)
      Move(in := 100, out1 => #Output)
   END_RUNG
   // the same network as SCL:
   IF "Expected/Value_All".V = "Expected/Value_All".Expected_81 THEN #Output := 81; END_IF;
   IF "Expected/Value_All".V = "Expected/Value_All".Expected_82 THEN #Output := 82; END_IF;
   IF "Expected/Value_All".V = "Expected/Value_All".Expected_83 THEN #Output := 83; END_IF;
   IF "Expected/Value_All".V = "Expected/Value_All".Expected_84 THEN #Output := 84; END_IF;
   IF "Expected/Value_All".V = "Expected/Value_All".Expected_85 THEN #Output := 85; END_IF;
   IF "Expected/Value_All".V = "Expected/Value_All".Expected_86 THEN #Output := 86; END_IF;
   IF "Expected/Value_All".V = "Expected/Value_All".Expected_87 THEN #Output := 87; END_IF;
   IF "Expected/Value_All".V = "Expected/Value_All".Expected_88 THEN #Output := 88; END_IF;
   IF "Expected/Value_All".V = "Expected/Value_All".Expected_89 THEN #Output := 89; END_IF;
   IF "Expected/Value_All".V = "Expected/Value_All".Expected_90 THEN #Output := 90; END_IF;
   IF "Expected/Value_All".V = "Expected/Value_All".Expected_91 THEN #Output := 91; END_IF;
   IF "Expected/Value_All".V = "Expected/Value_All".Expected_92 THEN #Output := 92; END_IF;
   IF "Expected/Value_All".V = "Expected/Value_All".Expected_93 THEN #Output := 93; END_IF;
   IF "Expected/Value_All".V = "Expected/Value_All".Expected_94 THEN #Output := 94; END_IF;
   IF "Expected/Value_All".V = "Expected/Value_All".Expected_95 THEN #Output := 95; END_IF;
   IF "Expected/Value_All".V = "Expected/Value_All".Expected_96 THEN #Output := 96; END_IF;
   IF "Expected/Value_All".V = "Expected/Value_All".Expected_97 THEN #Output := 97; END_IF;
   IF "Expected/Value_All".V = "Expected/Value_All".Expected_98 THEN #Output := 98; END_IF;
   IF "Expected/Value_All".V = "Expected/Value_All".Expected_99 THEN #Output := 99; END_IF;
   IF "Expected/Value_All".V = "Expected/Value_All".Expected_100 THEN #Output := 100; END_IF;
END_REGION

REGION Network 6
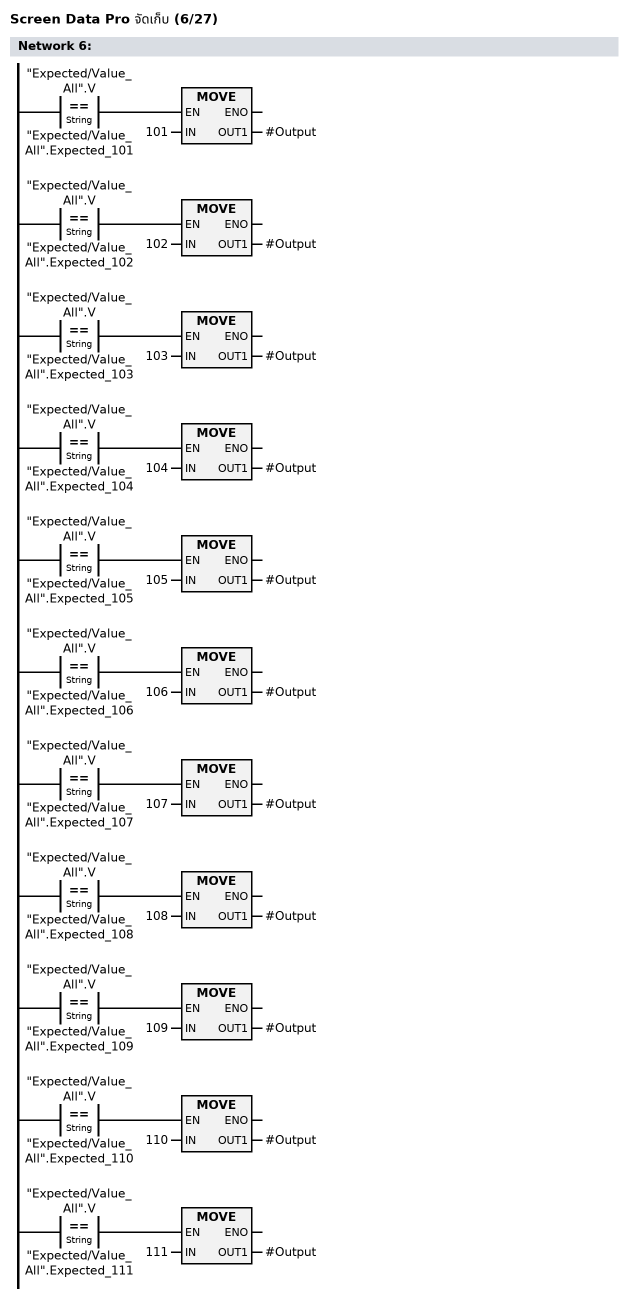
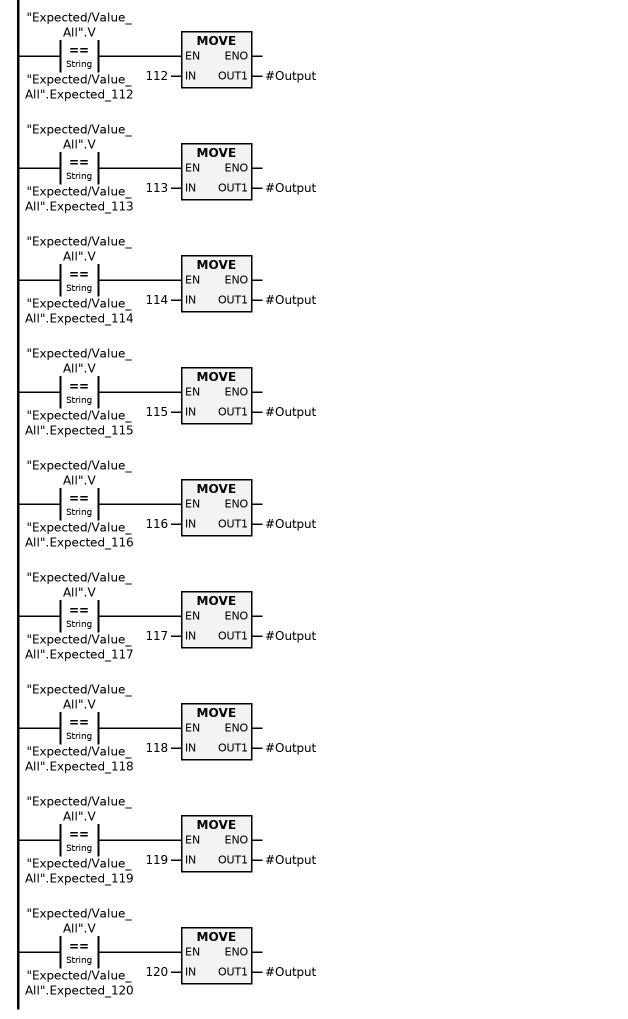
   RUNG wire#powerrail
      { S7_Templates := "SrcType := String" } EQ_Contact(in1 := "Expected/Value_All".V, in2 := "Expected/Value_All".Expected_101)
      Move(in := 101, out1 => #Output)
   END_RUNG
   RUNG wire#powerrail
      { S7_Templates := "SrcType := String" } EQ_Contact(in1 := "Expected/Value_All".V, in2 := "Expected/Value_All".Expected_102)
      Move(in := 102, out1 => #Output)
   END_RUNG
   RUNG wire#powerrail
      { S7_Templates := "SrcType := String" } EQ_Contact(in1 := "Expected/Value_All".V, in2 := "Expected/Value_All".Expected_103)
      Move(in := 103, out1 => #Output)
   END_RUNG
   RUNG wire#powerrail
      { S7_Templates := "SrcType := String" } EQ_Contact(in1 := "Expected/Value_All".V, in2 := "Expected/Value_All".Expected_104)
      Move(in := 104, out1 => #Output)
   END_RUNG
   RUNG wire#powerrail
      { S7_Templates := "SrcType := String" } EQ_Contact(in1 := "Expected/Value_All".V, in2 := "Expected/Value_All".Expected_105)
      Move(in := 105, out1 => #Output)
   END_RUNG
   RUNG wire#powerrail
      { S7_Templates := "SrcType := String" } EQ_Contact(in1 := "Expected/Value_All".V, in2 := "Expected/Value_All".Expected_106)
      Move(in := 106, out1 => #Output)
   END_RUNG
   RUNG wire#powerrail
      { S7_Templates := "SrcType := String" } EQ_Contact(in1 := "Expected/Value_All".V, in2 := "Expected/Value_All".Expected_107)
      Move(in := 107, out1 => #Output)
   END_RUNG
   RUNG wire#powerrail
      { S7_Templates := "SrcType := String" } EQ_Contact(in1 := "Expected/Value_All".V, in2 := "Expected/Value_All".Expected_108)
      Move(in := 108, out1 => #Output)
   END_RUNG
   RUNG wire#powerrail
      { S7_Templates := "SrcType := String" } EQ_Contact(in1 := "Expected/Value_All".V, in2 := "Expected/Value_All".Expected_109)
      Move(in := 109, out1 => #Output)
   END_RUNG
   RUNG wire#powerrail
      { S7_Templates := "SrcType := String" } EQ_Contact(in1 := "Expected/Value_All".V, in2 := "Expected/Value_All".Expected_110)
      Move(in := 110, out1 => #Output)
   END_RUNG
   RUNG wire#powerrail
      { S7_Templates := "SrcType := String" } EQ_Contact(in1 := "Expected/Value_All".V, in2 := "Expected/Value_All".Expected_111)
      Move(in := 111, out1 => #Output)
   END_RUNG
   RUNG wire#powerrail
      { S7_Templates := "SrcType := String" } EQ_Contact(in1 := "Expected/Value_All".V, in2 := "Expected/Value_All".Expected_112)
      Move(in := 112, out1 => #Output)
   END_RUNG
   RUNG wire#powerrail
      { S7_Templates := "SrcType := String" } EQ_Contact(in1 := "Expected/Value_All".V, in2 := "Expected/Value_All".Expected_113)
      Move(in := 113, out1 => #Output)
   END_RUNG
   RUNG wire#powerrail
      { S7_Templates := "SrcType := String" } EQ_Contact(in1 := "Expected/Value_All".V, in2 := "Expected/Value_All".Expected_114)
      Move(in := 114, out1 => #Output)
   END_RUNG
   RUNG wire#powerrail
      { S7_Templates := "SrcType := String" } EQ_Contact(in1 := "Expected/Value_All".V, in2 := "Expected/Value_All".Expected_115)
      Move(in := 115, out1 => #Output)
   END_RUNG
   RUNG wire#powerrail
      { S7_Templates := "SrcType := String" } EQ_Contact(in1 := "Expected/Value_All".V, in2 := "Expected/Value_All".Expected_116)
      Move(in := 116, out1 => #Output)
   END_RUNG
   RUNG wire#powerrail
      { S7_Templates := "SrcType := String" } EQ_Contact(in1 := "Expected/Value_All".V, in2 := "Expected/Value_All".Expected_117)
      Move(in := 117, out1 => #Output)
   END_RUNG
   RUNG wire#powerrail
      { S7_Templates := "SrcType := String" } EQ_Contact(in1 := "Expected/Value_All".V, in2 := "Expected/Value_All".Expected_118)
      Move(in := 118, out1 => #Output)
   END_RUNG
   RUNG wire#powerrail
      { S7_Templates := "SrcType := String" } EQ_Contact(in1 := "Expected/Value_All".V, in2 := "Expected/Value_All".Expected_119)
      Move(in := 119, out1 => #Output)
   END_RUNG
   RUNG wire#powerrail
      { S7_Templates := "SrcType := String" } EQ_Contact(in1 := "Expected/Value_All".V, in2 := "Expected/Value_All".Expected_120)
      Move(in := 120, out1 => #Output)
   END_RUNG
   // the same network as SCL:
   IF "Expected/Value_All".V = "Expected/Value_All".Expected_101 THEN #Output := 101; END_IF;
   IF "Expected/Value_All".V = "Expected/Value_All".Expected_102 THEN #Output := 102; END_IF;
   IF "Expected/Value_All".V = "Expected/Value_All".Expected_103 THEN #Output := 103; END_IF;
   IF "Expected/Value_All".V = "Expected/Value_All".Expected_104 THEN #Output := 104; END_IF;
   IF "Expected/Value_All".V = "Expected/Value_All".Expected_105 THEN #Output := 105; END_IF;
   IF "Expected/Value_All".V = "Expected/Value_All".Expected_106 THEN #Output := 106; END_IF;
   IF "Expected/Value_All".V = "Expected/Value_All".Expected_107 THEN #Output := 107; END_IF;
   IF "Expected/Value_All".V = "Expected/Value_All".Expected_108 THEN #Output := 108; END_IF;
   IF "Expected/Value_All".V = "Expected/Value_All".Expected_109 THEN #Output := 109; END_IF;
   IF "Expected/Value_All".V = "Expected/Value_All".Expected_110 THEN #Output := 110; END_IF;
   IF "Expected/Value_All".V = "Expected/Value_All".Expected_111 THEN #Output := 111; END_IF;
   IF "Expected/Value_All".V = "Expected/Value_All".Expected_112 THEN #Output := 112; END_IF;
   IF "Expected/Value_All".V = "Expected/Value_All".Expected_113 THEN #Output := 113; END_IF;
   IF "Expected/Value_All".V = "Expected/Value_All".Expected_114 THEN #Output := 114; END_IF;
   IF "Expected/Value_All".V = "Expected/Value_All".Expected_115 THEN #Output := 115; END_IF;
   IF "Expected/Value_All".V = "Expected/Value_All".Expected_116 THEN #Output := 116; END_IF;
   IF "Expected/Value_All".V = "Expected/Value_All".Expected_117 THEN #Output := 117; END_IF;
   IF "Expected/Value_All".V = "Expected/Value_All".Expected_118 THEN #Output := 118; END_IF;
   IF "Expected/Value_All".V = "Expected/Value_All".Expected_119 THEN #Output := 119; END_IF;
   IF "Expected/Value_All".V = "Expected/Value_All".Expected_120 THEN #Output := 120; END_IF;
END_REGION

REGION Network 7
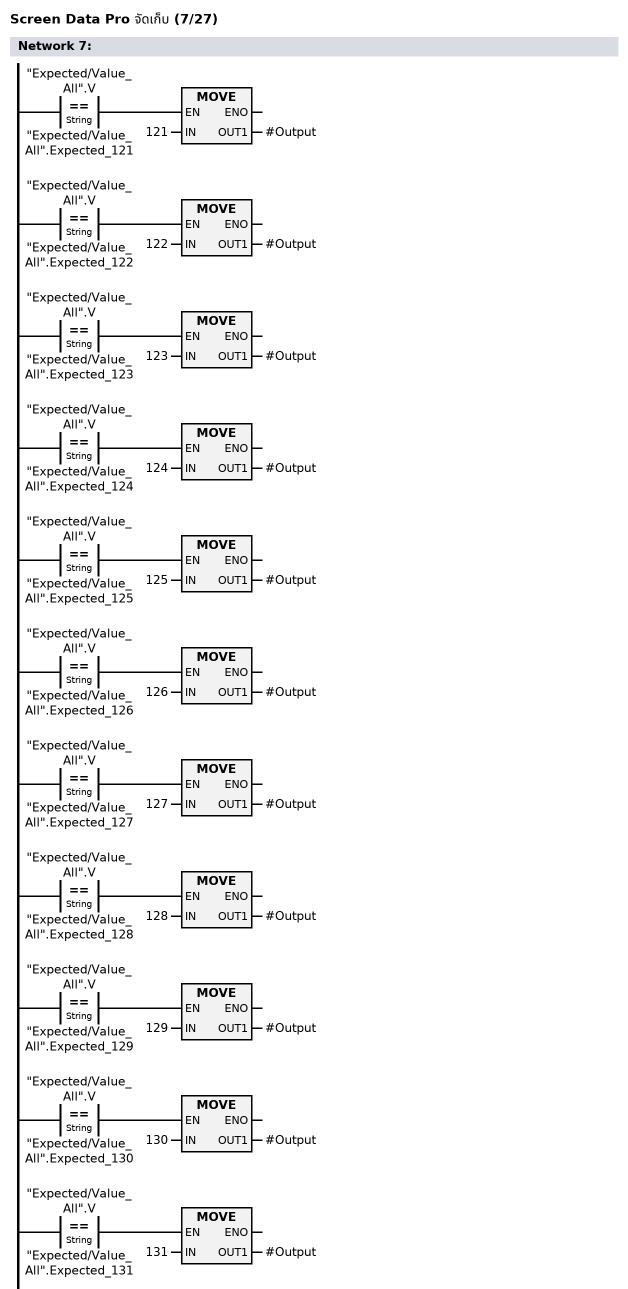
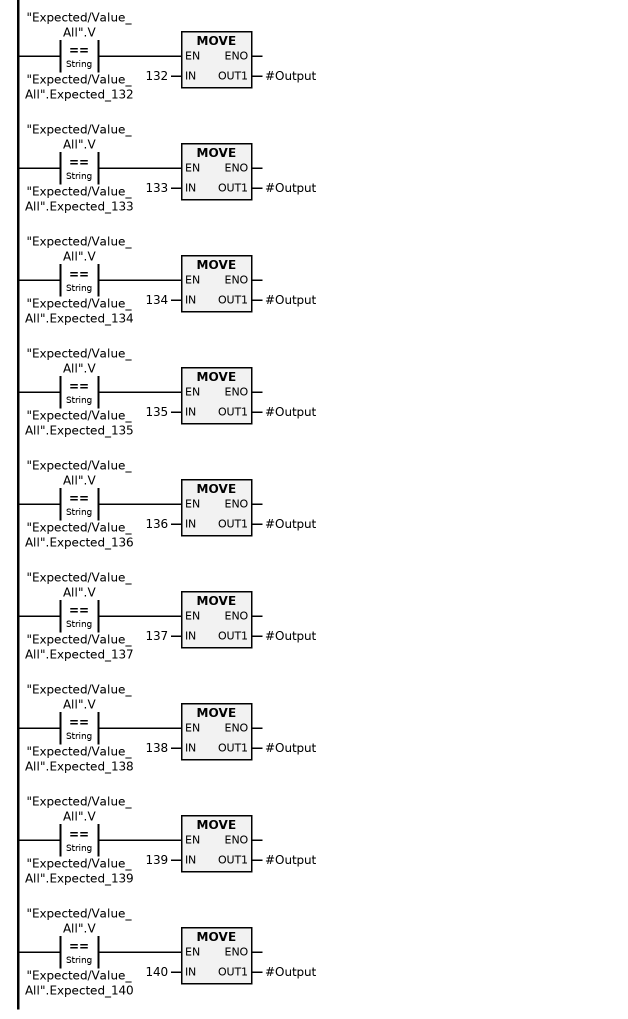
   RUNG wire#powerrail
      { S7_Templates := "SrcType := String" } EQ_Contact(in1 := "Expected/Value_All".V, in2 := "Expected/Value_All".Expected_121)
      Move(in := 121, out1 => #Output)
   END_RUNG
   RUNG wire#powerrail
      { S7_Templates := "SrcType := String" } EQ_Contact(in1 := "Expected/Value_All".V, in2 := "Expected/Value_All".Expected_122)
      Move(in := 122, out1 => #Output)
   END_RUNG
   RUNG wire#powerrail
      { S7_Templates := "SrcType := String" } EQ_Contact(in1 := "Expected/Value_All".V, in2 := "Expected/Value_All".Expected_123)
      Move(in := 123, out1 => #Output)
   END_RUNG
   RUNG wire#powerrail
      { S7_Templates := "SrcType := String" } EQ_Contact(in1 := "Expected/Value_All".V, in2 := "Expected/Value_All".Expected_124)
      Move(in := 124, out1 => #Output)
   END_RUNG
   RUNG wire#powerrail
      { S7_Templates := "SrcType := String" } EQ_Contact(in1 := "Expected/Value_All".V, in2 := "Expected/Value_All".Expected_125)
      Move(in := 125, out1 => #Output)
   END_RUNG
   RUNG wire#powerrail
      { S7_Templates := "SrcType := String" } EQ_Contact(in1 := "Expected/Value_All".V, in2 := "Expected/Value_All".Expected_126)
      Move(in := 126, out1 => #Output)
   END_RUNG
   RUNG wire#powerrail
      { S7_Templates := "SrcType := String" } EQ_Contact(in1 := "Expected/Value_All".V, in2 := "Expected/Value_All".Expected_127)
      Move(in := 127, out1 => #Output)
   END_RUNG
   RUNG wire#powerrail
      { S7_Templates := "SrcType := String" } EQ_Contact(in1 := "Expected/Value_All".V, in2 := "Expected/Value_All".Expected_128)
      Move(in := 128, out1 => #Output)
   END_RUNG
   RUNG wire#powerrail
      { S7_Templates := "SrcType := String" } EQ_Contact(in1 := "Expected/Value_All".V, in2 := "Expected/Value_All".Expected_129)
      Move(in := 129, out1 => #Output)
   END_RUNG
   RUNG wire#powerrail
      { S7_Templates := "SrcType := String" } EQ_Contact(in1 := "Expected/Value_All".V, in2 := "Expected/Value_All".Expected_130)
      Move(in := 130, out1 => #Output)
   END_RUNG
   RUNG wire#powerrail
      { S7_Templates := "SrcType := String" } EQ_Contact(in1 := "Expected/Value_All".V, in2 := "Expected/Value_All".Expected_131)
      Move(in := 131, out1 => #Output)
   END_RUNG
   RUNG wire#powerrail
      { S7_Templates := "SrcType := String" } EQ_Contact(in1 := "Expected/Value_All".V, in2 := "Expected/Value_All".Expected_132)
      Move(in := 132, out1 => #Output)
   END_RUNG
   RUNG wire#powerrail
      { S7_Templates := "SrcType := String" } EQ_Contact(in1 := "Expected/Value_All".V, in2 := "Expected/Value_All".Expected_133)
      Move(in := 133, out1 => #Output)
   END_RUNG
   RUNG wire#powerrail
      { S7_Templates := "SrcType := String" } EQ_Contact(in1 := "Expected/Value_All".V, in2 := "Expected/Value_All".Expected_134)
      Move(in := 134, out1 => #Output)
   END_RUNG
   RUNG wire#powerrail
      { S7_Templates := "SrcType := String" } EQ_Contact(in1 := "Expected/Value_All".V, in2 := "Expected/Value_All".Expected_135)
      Move(in := 135, out1 => #Output)
   END_RUNG
   RUNG wire#powerrail
      { S7_Templates := "SrcType := String" } EQ_Contact(in1 := "Expected/Value_All".V, in2 := "Expected/Value_All".Expected_136)
      Move(in := 136, out1 => #Output)
   END_RUNG
   RUNG wire#powerrail
      { S7_Templates := "SrcType := String" } EQ_Contact(in1 := "Expected/Value_All".V, in2 := "Expected/Value_All".Expected_137)
      Move(in := 137, out1 => #Output)
   END_RUNG
   RUNG wire#powerrail
      { S7_Templates := "SrcType := String" } EQ_Contact(in1 := "Expected/Value_All".V, in2 := "Expected/Value_All".Expected_138)
      Move(in := 138, out1 => #Output)
   END_RUNG
   RUNG wire#powerrail
      { S7_Templates := "SrcType := String" } EQ_Contact(in1 := "Expected/Value_All".V, in2 := "Expected/Value_All".Expected_139)
      Move(in := 139, out1 => #Output)
   END_RUNG
   RUNG wire#powerrail
      { S7_Templates := "SrcType := String" } EQ_Contact(in1 := "Expected/Value_All".V, in2 := "Expected/Value_All".Expected_140)
      Move(in := 140, out1 => #Output)
   END_RUNG
   // the same network as SCL:
   IF "Expected/Value_All".V = "Expected/Value_All".Expected_121 THEN #Output := 121; END_IF;
   IF "Expected/Value_All".V = "Expected/Value_All".Expected_122 THEN #Output := 122; END_IF;
   IF "Expected/Value_All".V = "Expected/Value_All".Expected_123 THEN #Output := 123; END_IF;
   IF "Expected/Value_All".V = "Expected/Value_All".Expected_124 THEN #Output := 124; END_IF;
   IF "Expected/Value_All".V = "Expected/Value_All".Expected_125 THEN #Output := 125; END_IF;
   IF "Expected/Value_All".V = "Expected/Value_All".Expected_126 THEN #Output := 126; END_IF;
   IF "Expected/Value_All".V = "Expected/Value_All".Expected_127 THEN #Output := 127; END_IF;
   IF "Expected/Value_All".V = "Expected/Value_All".Expected_128 THEN #Output := 128; END_IF;
   IF "Expected/Value_All".V = "Expected/Value_All".Expected_129 THEN #Output := 129; END_IF;
   IF "Expected/Value_All".V = "Expected/Value_All".Expected_130 THEN #Output := 130; END_IF;
   IF "Expected/Value_All".V = "Expected/Value_All".Expected_131 THEN #Output := 131; END_IF;
   IF "Expected/Value_All".V = "Expected/Value_All".Expected_132 THEN #Output := 132; END_IF;
   IF "Expected/Value_All".V = "Expected/Value_All".Expected_133 THEN #Output := 133; END_IF;
   IF "Expected/Value_All".V = "Expected/Value_All".Expected_134 THEN #Output := 134; END_IF;
   IF "Expected/Value_All".V = "Expected/Value_All".Expected_135 THEN #Output := 135; END_IF;
   IF "Expected/Value_All".V = "Expected/Value_All".Expected_136 THEN #Output := 136; END_IF;
   IF "Expected/Value_All".V = "Expected/Value_All".Expected_137 THEN #Output := 137; END_IF;
   IF "Expected/Value_All".V = "Expected/Value_All".Expected_138 THEN #Output := 138; END_IF;
   IF "Expected/Value_All".V = "Expected/Value_All".Expected_139 THEN #Output := 139; END_IF;
   IF "Expected/Value_All".V = "Expected/Value_All".Expected_140 THEN #Output := 140; END_IF;
END_REGION

REGION Network 8
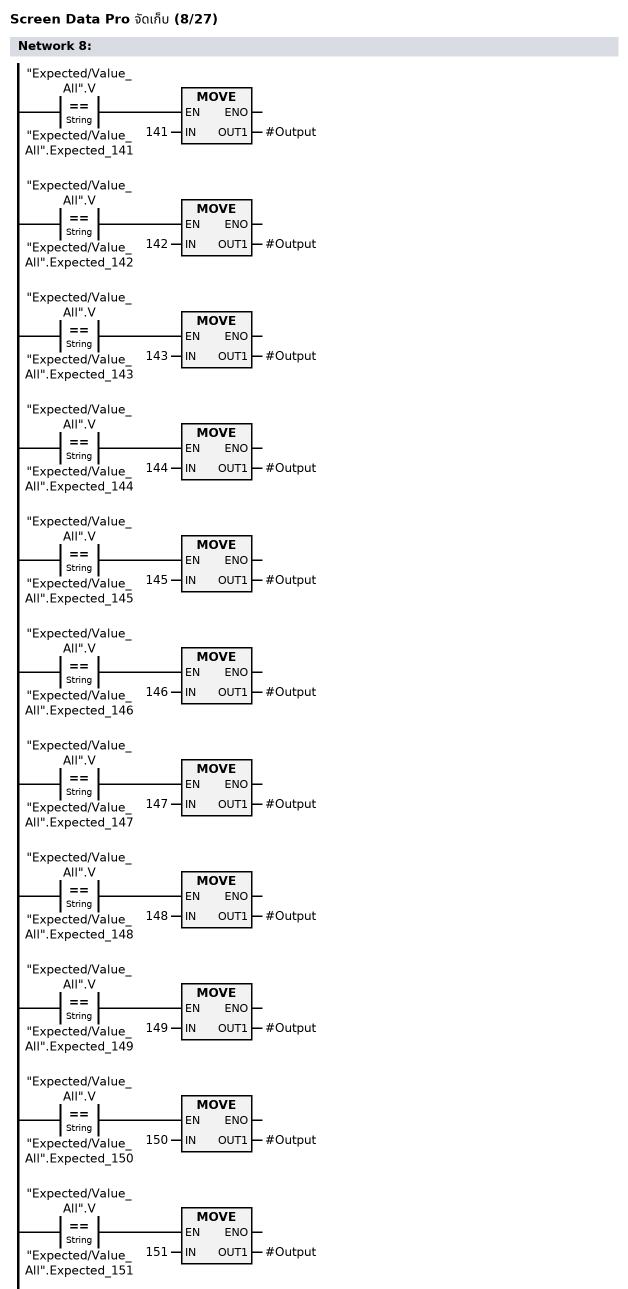
